screen "D_GraphicView_1" 800x480
   GraphicView "Static" at 6,4 size 100x60
   TextField "Label_Static" at 6,96 size 44x17; Text 'Static'
   GraphicView "A_Range" at 158,4 size 100x60
      Appearance <- "D_Range"
   TextField "Label_A_Range" at 158,96 size 63x17; Text 'A_Range'
   GraphicView "A_Flash" at 310,4 size 100x60
      Appearance <- "D_Range"
   TextField "Label_A_Flash" at 310,96 size 56x17; Text 'A_Flash'
   GraphicView "A_Bit" at 462,4 size 100x60
      Appearance <- "D_Bool"
   TextField "Label_A_Bit" at 462,96 size 40x17; Text 'A_Bit'
   GraphicView "A_Bits" at 614,4 size 100x60
      Appearance <- "D_Bits"
   TextField "Label_A_Bits" at 614,96 size 47x17; Text 'A_Bits'
   GraphicView "V_Range" at 6,116 size 100x60
      Visibility <- "D_Range"
   TextField "Label_V_Range" at 6,208 size 62x17; Text 'V_Range'
   GraphicView "V_Bit" at 158,116 size 100x60
      Visibility <- "D_Vis"
   TextField "Label_V_Bit" at 158,208 size 39x17; Text 'V_Bit'
   GraphicView "M_H" at 310,116 size 100x60
      HorizontalMovement <- "D_Pct"
   TextField "Label_M_H" at 310,208 size 33x17; Text 'M_H'
   GraphicView "M_V" at 462,116 size 100x60
      VerticalMovement <- "D_Pct"
   TextField "Label_M_V" at 462,208 size 32x17; Text 'M_V'
   GraphicView "M_D" at 614,116 size 100x60
      DiagonalMovement <- "D_Pct"
   TextField "Label_M_D" at 614,208 size 33x17; Text 'M_D'
   GraphicView "M_Direct" at 6,228 size 100x60
      DirectMovement <- "D_X"
      DirectMovement <- "D_Y"
   TextField "Label_M_Direct" at 6,320 size 64x17; Text 'M_Direct'
   GraphicView "E_Range" at 158,228 size 100x60
      ObjectEnable <- "D_Range"
   TextField "Label_E_Range" at 158,320 size 61x17; Text 'E_Range'
   GraphicView "E_Bit" at 310,228 size 100x60
      ObjectEnable <- "D_En"
   TextField "Label_E_Bit" at 310,320 size 38x17; Text 'E_Bit'
   IOField "State" at 4,454 size 60x22; FormatPattern 9
      ProcessValue <- "D_State"
   Button "S1" at 70,454 size 40x22; TextOff 'S1'
      on Click: "SetS1"()
   Button "S2" at 114,454 size 40x22; TextOff 'S2'
      on Click: "SetS2"()
   Button "S3" at 158,454 size 40x22; TextOff 'S3'
      on Click: "SetS3"()
   Button "S4" at 202,454 size 40x22; TextOff 'S4'
      on Click: "SetS4"()
   Button "Next" at 756,454 size 40x22; TextOff 'Next'
      on Click: ActivateScreen("D_IOField_1", 0)

screen "D_IOField_2" 800x480
   IOField "PV_Int_Output" at 6,4 size 100x30; FormatPattern s99999
      ProcessValue <- "D_Int"
   TextField "Label_PV_Int_Output" at 6,66 size 102x17; Text 'PV_Int_Output'
   IOField "PV_Int_s99" at 158,4 size 100x30; FormatPattern s99
      ProcessValue <- "D_Int"
   TextField "Label_PV_Int_s99" at 158,66 size 80x17; Text 'PV_Int_s99'
   IOField "State" at 4,454 size 60x22; FormatPattern 9
      ProcessValue <- "D_State"
   Button "S1" at 70,454 size 40x22; TextOff 'S1'
      on Click: "SetS1"()
   Button "S2" at 114,454 size 40x22; TextOff 'S2'
      on Click: "SetS2"()
   Button "S3" at 158,454 size 40x22; TextOff 'S3'
      on Click: "SetS3"()
   Button "S4" at 202,454 size 40x22; TextOff 'S4'
      on Click: "SetS4"()
   Button "Next" at 756,454 size 40x22; TextOff 'Next'
      on Click: ActivateScreen("D_Button_1", 0)

screen "D_Line_1" 800x480
   TextField "Label_Static" at 6,86 size 44x17; Text 'Static'
   Line "A_Range" at 158,4 size 100x50
      Appearance <- "D_Range"
   TextField "Label_A_Range" at 158,86 size 63x17; Text 'A_Range'
   Line "A_Flash" at 310,4 size 100x50
      Appearance <- "D_Range"
   TextField "Label_A_Flash" at 310,86 size 56x17; Text 'A_Flash'
   Line "A_Bit" at 462,4 size 100x50
      Appearance <- "D_Bool"
   TextField "Label_A_Bit" at 462,86 size 40x17; Text 'A_Bit'
   Line "A_Bits" at 614,4 size 100x50
      Appearance <- "D_Bits"
   TextField "Label_A_Bits" at 614,86 size 47x17; Text 'A_Bits'
   Line "V_Range" at 6,106 size 100x50
      Visibility <- "D_Range"
   TextField "Label_V_Range" at 6,188 size 62x17; Text 'V_Range'
   Line "V_Bit" at 158,106 size 100x50
      Visibility <- "D_Vis"
   TextField "Label_V_Bit" at 158,188 size 39x17; Text 'V_Bit'
   Line "M_H" at 310,106 size 100x50
      HorizontalMovement <- "D_Pct"
   TextField "Label_M_H" at 310,188 size 33x17; Text 'M_H'
   Line "M_V" at 462,106 size 100x50
      VerticalMovement <- "D_Pct"
   TextField "Label_M_V" at 462,188 size 32x17; Text 'M_V'
   Line "M_D" at 614,106 size 100x50
      DiagonalMovement <- "D_Pct"
   TextField "Label_M_D" at 614,188 size 33x17; Text 'M_D'
   Line "M_Direct" at 6,208 size 100x50
      DirectMovement <- "D_X"
      DirectMovement <- "D_Y"
   TextField "Label_M_Direct" at 6,290 size 64x17; Text 'M_Direct'
   Line "E_Range" at 158,208 size 100x50
      ObjectEnable <- "D_Range"
   TextField "Label_E_Range" at 158,290 size 61x17; Text 'E_Range'
   Line "E_Bit" at 310,208 size 100x50
      ObjectEnable <- "D_En"
   TextField "Label_E_Bit" at 310,290 size 38x17; Text 'E_Bit'
   IOField "State" at 4,454 size 60x22; FormatPattern 9
      ProcessValue <- "D_State"
   Button "S1" at 70,454 size 40x22; TextOff 'S1'
      on Click: "SetS1"()
   Button "S2" at 114,454 size 40x22; TextOff 'S2'
      on Click: "SetS2"()
   Button "S3" at 158,454 size 40x22; TextOff 'S3'
      on Click: "SetS3"()
   Button "S4" at 202,454 size 40x22; TextOff 'S4'
      on Click: "SetS4"()
   Button "Next" at 756,454 size 40x22; TextOff 'Next'
      on Click: ActivateScreen("D_Polyline_1", 0)

screen "D_Polygon_1" 800x480
   TextField "Label_Static" at 6,86 size 44x17; Text 'Static'
   Polygon "A_Range" at 158,4 size 100x50
      Appearance <- "D_Range"
   TextField "Label_A_Range" at 158,86 size 63x17; Text 'A_Range'
   Polygon "A_Flash" at 310,4 size 100x50
      Appearance <- "D_Range"
   TextField "Label_A_Flash" at 310,86 size 56x17; Text 'A_Flash'
   Polygon "A_Bit" at 462,4 size 100x50
      Appearance <- "D_Bool"
   TextField "Label_A_Bit" at 462,86 size 40x17; Text 'A_Bit'
   Polygon "A_Bits" at 614,4 size 100x50
      Appearance <- "D_Bits"
   TextField "Label_A_Bits" at 614,86 size 47x17; Text 'A_Bits'
   Polygon "V_Range" at 6,106 size 100x50
      Visibility <- "D_Range"
   TextField "Label_V_Range" at 6,188 size 62x17; Text 'V_Range'
   Polygon "V_Bit" at 158,106 size 100x50
      Visibility <- "D_Vis"
   TextField "Label_V_Bit" at 158,188 size 39x17; Text 'V_Bit'
   Polygon "M_H" at 310,106 size 100x50
      HorizontalMovement <- "D_Pct"
   TextField "Label_M_H" at 310,188 size 33x17; Text 'M_H'
   Polygon "M_V" at 462,106 size 100x50
      VerticalMovement <- "D_Pct"
   TextField "Label_M_V" at 462,188 size 32x17; Text 'M_V'
   Polygon "M_D" at 614,106 size 100x50
      DiagonalMovement <- "D_Pct"
   TextField "Label_M_D" at 614,188 size 33x17; Text 'M_D'
   Polygon "M_Direct" at 6,208 size 100x50
      DirectMovement <- "D_X"
      DirectMovement <- "D_Y"
   TextField "Label_M_Direct" at 6,290 size 64x17; Text 'M_Direct'
   Polygon "E_Range" at 158,208 size 100x50
      ObjectEnable <- "D_Range"
   TextField "Label_E_Range" at 158,290 size 61x17; Text 'E_Range'
   Polygon "E_Bit" at 310,208 size 100x50
      ObjectEnable <- "D_En"
   TextField "Label_E_Bit" at 310,290 size 38x17; Text 'E_Bit'
   IOField "State" at 4,454 size 60x22; FormatPattern 9
      ProcessValue <- "D_State"
   Button "S1" at 70,454 size 40x22; TextOff 'S1'
      on Click: "SetS1"()
   Button "S2" at 114,454 size 40x22; TextOff 'S2'
      on Click: "SetS2"()
   Button "S3" at 158,454 size 40x22; TextOff 'S3'
      on Click: "SetS3"()
   Button "S4" at 202,454 size 40x22; TextOff 'S4'
      on Click: "SetS4"()
   Button "Next" at 756,454 size 40x22; TextOff 'Next'
      on Click: ActivateScreen("D_Ellipse_1", 0)

screen "D_Polyline_1" 800x480
   TextField "Label_Static" at 6,86 size 44x17; Text 'Static'
   Polyline "A_Range" at 158,4 size 100x50
      Appearance <- "D_Range"
   TextField "Label_A_Range" at 158,86 size 63x17; Text 'A_Range'
   Polyline "A_Flash" at 310,4 size 100x50
      Appearance <- "D_Range"
   TextField "Label_A_Flash" at 310,86 size 56x17; Text 'A_Flash'
   Polyline "A_Bit" at 462,4 size 100x50
      Appearance <- "D_Bool"
   TextField "Label_A_Bit" at 462,86 size 40x17; Text 'A_Bit'
   Polyline "A_Bits" at 614,4 size 100x50
      Appearance <- "D_Bits"
   TextField "Label_A_Bits" at 614,86 size 47x17; Text 'A_Bits'
   Polyline "V_Range" at 6,106 size 100x50
      Visibility <- "D_Range"
   TextField "Label_V_Range" at 6,188 size 62x17; Text 'V_Range'
   Polyline "V_Bit" at 158,106 size 100x50
      Visibility <- "D_Vis"
   TextField "Label_V_Bit" at 158,188 size 39x17; Text 'V_Bit'
   Polyline "M_H" at 310,106 size 100x50
      HorizontalMovement <- "D_Pct"
   TextField "Label_M_H" at 310,188 size 33x17; Text 'M_H'
   Polyline "M_V" at 462,106 size 100x50
      VerticalMovement <- "D_Pct"
   TextField "Label_M_V" at 462,188 size 32x17; Text 'M_V'
   Polyline "M_D" at 614,106 size 100x50
      DiagonalMovement <- "D_Pct"
   TextField "Label_M_D" at 614,188 size 33x17; Text 'M_D'
   Polyline "M_Direct" at 6,208 size 100x50
      DirectMovement <- "D_X"
      DirectMovement <- "D_Y"
   TextField "Label_M_Direct" at 6,290 size 64x17; Text 'M_Direct'
   Polyline "E_Range" at 158,208 size 100x50
      ObjectEnable <- "D_Range"
   TextField "Label_E_Range" at 158,290 size 61x17; Text 'E_Range'
   Polyline "E_Bit" at 310,208 size 100x50
      ObjectEnable <- "D_En"
   TextField "Label_E_Bit" at 310,290 size 38x17; Text 'E_Bit'
   IOField "State" at 4,454 size 60x22; FormatPattern 9
      ProcessValue <- "D_State"
   Button "S1" at 70,454 size 40x22; TextOff 'S1'
      on Click: "SetS1"()
   Button "S2" at 114,454 size 40x22; TextOff 'S2'
      on Click: "SetS2"()
   Button "S3" at 158,454 size 40x22; TextOff 'S3'
      on Click: "SetS3"()
   Button "S4" at 202,454 size 40x22; TextOff 'S4'
      on Click: "SetS4"()
   Button "Next" at 756,454 size 40x22; TextOff 'Next'
      on Click: ActivateScreen("D_Polygon_1", 0)

screen "D_Rectangle_1" 800x480
   TextField "Label_Static" at 6,86 size 44x17; Text 'Static'
   Rectangle "A_Range" at 158,4 size 100x50
      Appearance <- "D_Range"
   TextField "Label_A_Range" at 158,86 size 63x17; Text 'A_Range'
   Rectangle "A_Flash" at 310,4 size 100x50
      Appearance <- "D_Range"
   TextField "Label_A_Flash" at 310,86 size 56x17; Text 'A_Flash'
   Rectangle "A_Bit" at 462,4 size 100x50
      Appearance <- "D_Bool"
   TextField "Label_A_Bit" at 462,86 size 40x17; Text 'A_Bit'
   Rectangle "A_Bits" at 614,4 size 100x50
      Appearance <- "D_Bits"
   TextField "Label_A_Bits" at 614,86 size 47x17; Text 'A_Bits'
   Rectangle "V_Range" at 6,106 size 100x50
      Visibility <- "D_Range"
   TextField "Label_V_Range" at 6,188 size 62x17; Text 'V_Range'
   Rectangle "V_Bit" at 158,106 size 100x50
      Visibility <- "D_Vis"
   TextField "Label_V_Bit" at 158,188 size 39x17; Text 'V_Bit'
   Rectangle "M_H" at 310,106 size 100x50
      HorizontalMovement <- "D_Pct"
   TextField "Label_M_H" at 310,188 size 33x17; Text 'M_H'
   Rectangle "M_V" at 462,106 size 100x50
      VerticalMovement <- "D_Pct"
   TextField "Label_M_V" at 462,188 size 32x17; Text 'M_V'
   Rectangle "M_D" at 614,106 size 100x50
      DiagonalMovement <- "D_Pct"
   TextField "Label_M_D" at 614,188 size 33x17; Text 'M_D'
   Rectangle "M_Direct" at 6,208 size 100x50
      DirectMovement <- "D_X"
      DirectMovement <- "D_Y"
   TextField "Label_M_Direct" at 6,290 size 64x17; Text 'M_Direct'
   Rectangle "E_Range" at 158,208 size 100x50
      ObjectEnable <- "D_Range"
   TextField "Label_E_Range" at 158,290 size 61x17; Text 'E_Range'
   Rectangle "E_Bit" at 310,208 size 100x50
      ObjectEnable <- "D_En"
   TextField "Label_E_Bit" at 310,290 size 38x17; Text 'E_Bit'
   IOField "State" at 4,454 size 60x22; FormatPattern 9
      ProcessValue <- "D_State"
   Button "S1" at 70,454 size 40x22; TextOff 'S1'
      on Click: "SetS1"()
   Button "S2" at 114,454 size 40x22; TextOff 'S2'
      on Click: "SetS2"()
   Button "S3" at 158,454 size 40x22; TextOff 'S3'
      on Click: "SetS3"()
   Button "S4" at 202,454 size 40x22; TextOff 'S4'
      on Click: "SetS4"()
   Button "Next" at 756,454 size 40x22; TextOff 'Next'
      on Click: ActivateScreen("D_TextField_1", 0)

screen "D_Switch_1" 800x480
   Switch "Static" at 6,4 size 120x40; CaptionText 'Switch'; TextOff '0'; TextOn '1'
   TextField "Label_Static" at 6,76 size 44x17; Text 'Static'
   Switch "A_Range" at 178,4 size 120x40; CaptionText 'Switch'; TextOff '0'; TextOn '1'
      Appearance <- "D_Range"
   TextField "Label_A_Range" at 178,76 size 63x17; Text 'A_Range'
   Switch "A_Flash" at 350,4 size 120x40; CaptionText 'Switch'; TextOff '0'; TextOn '1'
      Appearance <- "D_Range"
   TextField "Label_A_Flash" at 350,76 size 56x17; Text 'A_Flash'
   Switch "A_Bit" at 522,4 size 120x40; CaptionText 'Switch'; TextOff '0'; TextOn '1'
      Appearance <- "D_Bool"
   TextField "Label_A_Bit" at 522,76 size 40x17; Text 'A_Bit'
   Switch "A_Bits" at 6,96 size 120x40; CaptionText 'Switch'; TextOff '0'; TextOn '1'
      Appearance <- "D_Bits"
   TextField "Label_A_Bits" at 6,168 size 47x17; Text 'A_Bits'
   Switch "V_Range" at 178,96 size 120x40; CaptionText 'Switch'; TextOff '0'; TextOn '1'
      Visibility <- "D_Range"
   TextField "Label_V_Range" at 178,168 size 62x17; Text 'V_Range'
   Switch "V_Bit" at 350,96 size 120x40; CaptionText 'Switch'; TextOff '0'; TextOn '1'
      Visibility <- "D_Vis"
   TextField "Label_V_Bit" at 350,168 size 39x17; Text 'V_Bit'
   Switch "M_H" at 522,96 size 120x40; CaptionText 'Switch'; TextOff '0'; TextOn '1'
      HorizontalMovement <- "D_Pct"
   TextField "Label_M_H" at 522,168 size 33x17; Text 'M_H'
   Switch "M_V" at 6,188 size 120x40; CaptionText 'Switch'; TextOff '0'; TextOn '1'
      VerticalMovement <- "D_Pct"
   TextField "Label_M_V" at 6,260 size 32x17; Text 'M_V'
   Switch "M_D" at 178,188 size 120x40; CaptionText 'Switch'; TextOff '0'; TextOn '1'
      DiagonalMovement <- "D_Pct"
   TextField "Label_M_D" at 178,260 size 33x17; Text 'M_D'
   Switch "M_Direct" at 350,188 size 120x40; CaptionText 'Switch'; TextOff '0'; TextOn '1'
      DirectMovement <- "D_X"
      DirectMovement <- "D_Y"
   TextField "Label_M_Direct" at 350,260 size 64x17; Text 'M_Direct'
   Switch "E_Range" at 522,188 size 120x40; CaptionText 'Switch'; TextOff '0'; TextOn '1'
      ObjectEnable <- "D_Range"
   TextField "Label_E_Range" at 522,260 size 61x17; Text 'E_Range'
   Switch "E_Bit" at 6,280 size 120x40; CaptionText 'Switch'; TextOff '0'; TextOn '1'
      ObjectEnable <- "D_En"
   TextField "Label_E_Bit" at 6,352 size 38x17; Text 'E_Bit'
   Switch "PV_Bool" at 178,280 size 120x40; CaptionText 'Switch'; TextOff '0'; TextOn '1'
      ProcessValue <- "D_Bool"
   TextField "Label_PV_Bool" at 178,352 size 57x17; Text 'PV_Bool'
   IOField "State" at 4,454 size 60x22; FormatPattern 9
      ProcessValue <- "D_State"
   Button "S1" at 70,454 size 40x22; TextOff 'S1'
      on Click: "SetS1"()
   Button "S2" at 114,454 size 40x22; TextOff 'S2'
      on Click: "SetS2"()
   Button "S3" at 158,454 size 40x22; TextOff 'S3'
      on Click: "SetS3"()
   Button "S4" at 202,454 size 40x22; TextOff 'S4'
      on Click: "SetS4"()
   Button "Next" at 756,454 size 40x22; TextOff 'Next'
      on Click: ActivateScreen("D_SymbolLibrary_1", 0)

screen "D_SymbolicIOField_1" 800x480
   SymbolicIOField "Static" at 6,4 size 120x30; TextOff '0'; TextOn '1'
   TextField "Label_Static" at 6,66 size 44x17; Text 'Static'
   SymbolicIOField "A_Range" at 178,4 size 120x30; TextOff '0'; TextOn '1'
      Appearance <- "D_Range"
   TextField "Label_A_Range" at 178,66 size 63x17; Text 'A_Range'
   SymbolicIOField "A_Flash" at 350,4 size 120x30; TextOff '0'; TextOn '1'
      Appearance <- "D_Range"
   TextField "Label_A_Flash" at 350,66 size 56x17; Text 'A_Flash'
   SymbolicIOField "A_Bit" at 522,4 size 120x30; TextOff '0'; TextOn '1'
      Appearance <- "D_Bool"
   TextField "Label_A_Bit" at 522,66 size 40x17; Text 'A_Bit'
   SymbolicIOField "A_Bits" at 6,86 size 120x30; TextOff '0'; TextOn '1'
      Appearance <- "D_Bits"
   TextField "Label_A_Bits" at 6,148 size 47x17; Text 'A_Bits'
   SymbolicIOField "V_Range" at 178,86 size 120x30; TextOff '0'; TextOn '1'
      Visibility <- "D_Range"
   TextField "Label_V_Range" at 178,148 size 62x17; Text 'V_Range'
   SymbolicIOField "V_Bit" at 350,86 size 120x30; TextOff '0'; TextOn '1'
      Visibility <- "D_Vis"
   TextField "Label_V_Bit" at 350,148 size 39x17; Text 'V_Bit'
   SymbolicIOField "M_H" at 522,86 size 120x30; TextOff '0'; TextOn '1'
      HorizontalMovement <- "D_Pct"
   TextField "Label_M_H" at 522,148 size 33x17; Text 'M_H'
   SymbolicIOField "M_V" at 6,168 size 120x30; TextOff '0'; TextOn '1'
      VerticalMovement <- "D_Pct"
   TextField "Label_M_V" at 6,230 size 32x17; Text 'M_V'
   SymbolicIOField "M_D" at 178,168 size 120x30; TextOff '0'; TextOn '1'
      DiagonalMovement <- "D_Pct"
   TextField "Label_M_D" at 178,230 size 33x17; Text 'M_D'
   SymbolicIOField "M_Direct" at 350,168 size 120x30; TextOff '0'; TextOn '1'
      DirectMovement <- "D_X"
      DirectMovement <- "D_Y"
   TextField "Label_M_Direct" at 350,230 size 64x17; Text 'M_Direct'
   SymbolicIOField "E_Range" at 522,168 size 120x30; TextOff '0'; TextOn '1'
      ObjectEnable <- "D_Range"
   TextField "Label_E_Range" at 522,230 size 61x17; Text 'E_Range'
   SymbolicIOField "E_Bit" at 6,250 size 120x30; TextOff '0'; TextOn '1'
      ObjectEnable <- "D_En"
   TextField "Label_E_Bit" at 6,312 size 38x17; Text 'E_Bit'
   SymbolicIOField "PV_TL_Value" at 178,250 size 120x30; TextOff '0'; TextOn '1'; TextList "TL_Value"
      ProcessValue <- "D_TL"
   TextField "Label_PV_TL_Value" at 178,312 size 88x17; Text 'PV_TL_Value'
   SymbolicIOField "PV_TL_Bit" at 350,250 size 120x30; TextOff '0'; TextOn '1'; TextList "TL_Bit"
      ProcessValue <- "D_Bool"
   TextField "Label_PV_TL_Bit" at 350,312 size 70x17; Text 'PV_TL_Bit'
   SymbolicIOField "PV_TL_BitNo" at 522,250 size 120x30; TextOff '0'; TextOn '1'; TextList "TL_BitNo"
      ProcessValue <- "D_Bits"
   TextField "Label_PV_TL_BitNo" at 522,312 size 86x17; Text 'PV_TL_BitNo'
   IOField "State" at 4,454 size 60x22; FormatPattern 9
      ProcessValue <- "D_State"
   Button "S1" at 70,454 size 40x22; TextOff 'S1'
      on Click: "SetS1"()
   Button "S2" at 114,454 size 40x22; TextOff 'S2'
      on Click: "SetS2"()
   Button "S3" at 158,454 size 40x22; TextOff 'S3'
      on Click: "SetS3"()
   Button "S4" at 202,454 size 40x22; TextOff 'S4'
      on Click: "SetS4"()
   Button "Next" at 756,454 size 40x22; TextOff 'Next'
      on Click: ActivateScreen("D_GraphicIOField_1", 0)

screen "D_TextField_1" 800x480
   TextField "Static" at 6,4 size 35x17; Text 'Text'
   TextField "Label_Static" at 6,66 size 44x17; Text 'Static'
   TextField "A_Range" at 158,4 size 35x17; Text 'Text'
      Appearance <- "D_Range"
   TextField "Label_A_Range" at 158,66 size 63x17; Text 'A_Range'
   TextField "A_Flash" at 310,4 size 35x17; Text 'Text'
      Appearance <- "D_Range"
   TextField "Label_A_Flash" at 310,66 size 56x17; Text 'A_Flash'
   TextField "A_Bit" at 462,4 size 35x17; Text 'Text'
      Appearance <- "D_Bool"
   TextField "Label_A_Bit" at 462,66 size 40x17; Text 'A_Bit'
   TextField "A_Bits" at 614,4 size 35x17; Text 'Text'
      Appearance <- "D_Bits"
   TextField "Label_A_Bits" at 614,66 size 47x17; Text 'A_Bits'
   TextField "V_Range" at 6,86 size 35x17; Text 'Text'
      Visibility <- "D_Range"
   TextField "Label_V_Range" at 6,148 size 62x17; Text 'V_Range'
   TextField "V_Bit" at 158,86 size 35x17; Text 'Text'
      Visibility <- "D_Vis"
   TextField "Label_V_Bit" at 158,148 size 39x17; Text 'V_Bit'
   TextField "M_H" at 310,86 size 35x17; Text 'Text'
      HorizontalMovement <- "D_Pct"
   TextField "Label_M_H" at 310,148 size 33x17; Text 'M_H'
   TextField "M_V" at 462,86 size 35x17; Text 'Text'
      VerticalMovement <- "D_Pct"
   TextField "Label_M_V" at 462,148 size 32x17; Text 'M_V'
   TextField "M_D" at 614,86 size 35x17; Text 'Text'
      DiagonalMovement <- "D_Pct"
   TextField "Label_M_D" at 614,148 size 33x17; Text 'M_D'
   TextField "M_Direct" at 6,168 size 35x17; Text 'Text'
      DirectMovement <- "D_X"
      DirectMovement <- "D_Y"
   TextField "Label_M_Direct" at 6,230 size 64x17; Text 'M_Direct'
   TextField "E_Range" at 158,168 size 35x17; Text 'Text'
      ObjectEnable <- "D_Range"
   TextField "Label_E_Range" at 158,230 size 61x17; Text 'E_Range'
   TextField "E_Bit" at 310,168 size 35x17; Text 'Text'
      ObjectEnable <- "D_En"
   TextField "Label_E_Bit" at 310,230 size 38x17; Text 'E_Bit'
   IOField "State" at 4,454 size 60x22; FormatPattern 9
      ProcessValue <- "D_State"
   Button "S1" at 70,454 size 40x22; TextOff 'S1'
      on Click: "SetS1"()
   Button "S2" at 114,454 size 40x22; TextOff 'S2'
      on Click: "SetS2"()
   Button "S3" at 158,454 size 40x22; TextOff 'S3'
      on Click: "SetS3"()
   Button "S4" at 202,454 size 40x22; TextOff 'S4'
      on Click: "SetS4"()
   Button "Next" at 756,454 size 40x22; TextOff 'Next'
      on Click: ActivateScreen("D_GraphicView_1", 0)

screen "D_IOField_1" 800x480
   IOField "Static" at 6,4 size 100x30
   TextField "Label_Static" at 6,66 size 44x17; Text 'Static'
   IOField "A_Range" at 158,4 size 100x30
      Appearance <- "D_Range"
   TextField "Label_A_Range" at 158,66 size 63x17; Text 'A_Range'
   IOField "A_Flash" at 310,4 size 100x30
      Appearance <- "D_Range"
   TextField "Label_A_Flash" at 310,66 size 56x17; Text 'A_Flash'
   IOField "A_Bit" at 462,4 size 100x30
      Appearance <- "D_Bool"
   TextField "Label_A_Bit" at 462,66 size 40x17; Text 'A_Bit'
   IOField "A_Bits" at 614,4 size 100x30
      Appearance <- "D_Bits"
   TextField "Label_A_Bits" at 614,66 size 47x17; Text 'A_Bits'
   IOField "V_Range" at 6,86 size 100x30
      Visibility <- "D_Range"
   TextField "Label_V_Range" at 6,148 size 62x17; Text 'V_Range'
   IOField "V_Bit" at 158,86 size 100x30
      Visibility <- "D_Vis"
   TextField "Label_V_Bit" at 158,148 size 39x17; Text 'V_Bit'
   IOField "M_H" at 310,86 size 100x30
      HorizontalMovement <- "D_Pct"
   TextField "Label_M_H" at 310,148 size 33x17; Text 'M_H'
   IOField "M_V" at 462,86 size 100x30
      VerticalMovement <- "D_Pct"
   TextField "Label_M_V" at 462,148 size 32x17; Text 'M_V'
   IOField "M_D" at 614,86 size 100x30
      DiagonalMovement <- "D_Pct"
   TextField "Label_M_D" at 614,148 size 33x17; Text 'M_D'
   IOField "M_Direct" at 6,168 size 100x30
      DirectMovement <- "D_X"
      DirectMovement <- "D_Y"
   TextField "Label_M_Direct" at 6,230 size 64x17; Text 'M_Direct'
   IOField "E_Range" at 158,168 size 100x30
      ObjectEnable <- "D_Range"
   TextField "Label_E_Range" at 158,230 size 61x17; Text 'E_Range'
   IOField "E_Bit" at 310,168 size 100x30
      ObjectEnable <- "D_En"
   TextField "Label_E_Bit" at 310,230 size 38x17; Text 'E_Bit'
   IOField "PV_SInt" at 462,168 size 100x30; FormatPattern s999
      ProcessValue <- "D_SInt"
   TextField "Label_PV_SInt" at 462,230 size 57x17; Text 'PV_SInt'
   IOField "PV_Int" at 614,168 size 100x30; FormatPattern s99999
      ProcessValue <- "D_Int"
   TextField "Label_PV_Int" at 614,230 size 49x17; Text 'PV_Int'
   IOField "PV_DInt" at 6,250 size 100x30; FormatPattern s9999999999
      ProcessValue <- "D_DInt"
   TextField "Label_PV_DInt" at 6,312 size 58x17; Text 'PV_DInt'
   IOField "PV_USInt" at 158,250 size 100x30; FormatPattern 999
      ProcessValue <- "D_USInt"
   TextField "Label_PV_USInt" at 158,312 size 66x17; Text 'PV_USInt'
   IOField "PV_UInt" at 310,250 size 100x30; FormatPattern 99999
      ProcessValue <- "D_UInt"
   TextField "Label_PV_UInt" at 310,312 size 58x17; Text 'PV_UInt'
   IOField "PV_UDInt" at 462,250 size 100x30; FormatPattern 9999999999
      ProcessValue <- "D_UDInt"
   TextField "Label_PV_UDInt" at 462,312 size 67x17; Text 'PV_UDInt'
   IOField "PV_Real" at 614,250 size 100x30
      ProcessValue <- "D_Real"
   TextField "Label_PV_Real" at 614,312 size 58x17; Text 'PV_Real'
   IOField "PV_LReal" at 6,332 size 100x30
      ProcessValue <- "D_LReal"
   TextField "Label_PV_LReal" at 6,394 size 65x17; Text 'PV_LReal'
   IOField "PV_String" at 158,332 size 100x30
      ProcessValue <- "D_String"
   TextField "Label_PV_String" at 158,394 size 69x17; Text 'PV_String'
   IOField "PV_Int_Shift2" at 310,332 size 100x30; FormatPattern s99999
      ProcessValue <- "D_Int"
   TextField "Label_PV_Int_Shift2" at 310,394 size 96x17; Text 'PV_Int_Shift2'
   IOField "PV_Int_s999999" at 462,332 size 100x30; FormatPattern s999999
      ProcessValue <- "D_Int"
   TextField "Label_PV_Int_s999999" at 462,394 size 112x17; Text 'PV_Int_s999999'
   IOField "PV_Real_s9999_99" at 614,332 size 100x30; FormatPattern s9999.99
      ProcessValue <- "D_Real"
   TextField "Label_PV_Real_s9999_99" at 614,394 size 129x17; Text 'PV_Real_s9999_99'
   IOField "State" at 4,454 size 60x22; FormatPattern 9
      ProcessValue <- "D_State"
   Button "S1" at 70,454 size 40x22; TextOff 'S1'
      on Click: "SetS1"()
   Button "S2" at 114,454 size 40x22; TextOff 'S2'
      on Click: "SetS2"()
   Button "S3" at 158,454 size 40x22; TextOff 'S3'
      on Click: "SetS3"()
   Button "S4" at 202,454 size 40x22; TextOff 'S4'
      on Click: "SetS4"()
   Button "Next" at 756,454 size 40x22; TextOff 'Next'
      on Click: ActivateScreen("D_IOField_2", 0)

screen "D_Bar_1" 800x480
   Bar "Static" at 6,4 size 40x120
   TextField "Label_Static" at 6,156 size 44x17; Text 'Static'
   Bar "A_Range" at 98,4 size 40x120
      Appearance <- "D_Range"
   TextField "Label_A_Range" at 98,156 size 63x17; Text 'A_Range'
   Bar "A_Flash" at 190,4 size 40x120
      Appearance <- "D_Range"
   TextField "Label_A_Flash" at 190,156 size 56x17; Text 'A_Flash'
   Bar "A_Bit" at 282,4 size 40x120
      Appearance <- "D_Bool"
   TextField "Label_A_Bit" at 282,156 size 40x17; Text 'A_Bit'
   Bar "A_Bits" at 374,4 size 40x120
      Appearance <- "D_Bits"
   TextField "Label_A_Bits" at 374,156 size 47x17; Text 'A_Bits'
   Bar "V_Range" at 466,4 size 40x120
      Visibility <- "D_Range"
   TextField "Label_V_Range" at 466,156 size 62x17; Text 'V_Range'
   Bar "V_Bit" at 558,4 size 40x120
      Visibility <- "D_Vis"
   TextField "Label_V_Bit" at 558,156 size 39x17; Text 'V_Bit'
   Bar "M_H" at 650,4 size 40x120
      HorizontalMovement <- "D_Pct"
   TextField "Label_M_H" at 650,156 size 33x17; Text 'M_H'
   Bar "M_V" at 6,176 size 40x120
      VerticalMovement <- "D_Pct"
   TextField "Label_M_V" at 6,328 size 32x17; Text 'M_V'
   Bar "M_D" at 98,176 size 40x120
      DiagonalMovement <- "D_Pct"
   TextField "Label_M_D" at 98,328 size 33x17; Text 'M_D'
   Bar "M_Direct" at 190,176 size 40x120
      DirectMovement <- "D_X"
      DirectMovement <- "D_Y"
   TextField "Label_M_Direct" at 190,328 size 64x17; Text 'M_Direct'
   Bar "E_Range" at 282,176 size 40x120
      ObjectEnable <- "D_Range"
   TextField "Label_E_Range" at 282,328 size 61x17; Text 'E_Range'
   Bar "E_Bit" at 374,176 size 40x120
      ObjectEnable <- "D_En"
   TextField "Label_E_Bit" at 374,328 size 38x17; Text 'E_Bit'
   Bar "PV_Pct" at 466,176 size 40x120
      ProcessValue <- "D_Pct"
   TextField "Label_PV_Pct" at 466,328 size 50x17; Text 'PV_Pct'
   Bar "PV_Real" at 558,176 size 40x120
      ProcessValue <- "D_Real"
   TextField "Label_PV_Real" at 558,328 size 58x17; Text 'PV_Real'
   Bar "PV_BarR" at 650,176 size 40x120
      ProcessValue <- "D_BarR"
   TextField "Label_PV_BarR" at 650,328 size 60x17; Text 'PV_BarR'
   IOField "State" at 4,454 size 60x22; FormatPattern 9
      ProcessValue <- "D_State"
   Button "S1" at 70,454 size 40x22; TextOff 'S1'
      on Click: "SetS1"()
   Button "S2" at 114,454 size 40x22; TextOff 'S2'
      on Click: "SetS2"()
   Button "S3" at 158,454 size 40x22; TextOff 'S3'
      on Click: "SetS3"()
   Button "S4" at 202,454 size 40x22; TextOff 'S4'
      on Click: "SetS4"()
   Button "Next" at 756,454 size 40x22; TextOff 'Next'
      on Click: ActivateScreen("D_Bar_2", 0)

screen "D_Bar_2" 800x480
   Bar "PV_Pct_0_100" at 6,4 size 40x120; MinimumValue 0; MaximumValue 100
      ProcessValue <- "D_Pct"
   TextField "Label_PV_Pct_0_100" at 6,156 size 98x17; Text 'PV_Pct_0_100'
   Bar "PV_Pct_MaxMin" at 98,4 size 40x120
      ProcessValue <- "D_Pct"
      MaximumValue <- "D_Max"
      MinimumValue <- "D_Min"
   TextField "Label_PV_Pct_MaxMin" at 98,156 size 108x17; Text 'PV_Pct_MaxMin'
   IOField "State" at 4,454 size 60x22; FormatPattern 9
      ProcessValue <- "D_State"
   Button "S1" at 70,454 size 40x22; TextOff 'S1'
      on Click: "SetS1"()
   Button "S2" at 114,454 size 40x22; TextOff 'S2'
      on Click: "SetS2"()
   Button "S3" at 158,454 size 40x22; TextOff 'S3'
      on Click: "SetS3"()
   Button "S4" at 202,454 size 40x22; TextOff 'S4'
      on Click: "SetS4"()
   Button "Next" at 756,454 size 40x22; TextOff 'Next'
      on Click: ActivateScreen("D_Switch_1", 0)

screen "D_Gauge_1" 800x480
   Gauge "Static" at 6,4 size 150x150; CaptionText 'SIMATIC'
   TextField "Label_Static" at 6,186 size 44x17; Text 'Static'
   Gauge "A_Range" at 208,4 size 150x150; CaptionText 'SIMATIC'
      Appearance <- "D_Range"
   TextField "Label_A_Range" at 208,186 size 63x17; Text 'A_Range'
   Gauge "A_Flash" at 410,4 size 150x150; CaptionText 'SIMATIC'
      Appearance <- "D_Range"
   TextField "Label_A_Flash" at 410,186 size 56x17; Text 'A_Flash'
   Gauge "A_Bit" at 6,206 size 150x150; CaptionText 'SIMATIC'
      Appearance <- "D_Bool"
   TextField "Label_A_Bit" at 6,388 size 40x17; Text 'A_Bit'
   Gauge "A_Bits" at 208,206 size 150x150; CaptionText 'SIMATIC'
      Appearance <- "D_Bits"
   TextField "Label_A_Bits" at 208,388 size 47x17; Text 'A_Bits'
   Gauge "V_Range" at 410,206 size 150x150; CaptionText 'SIMATIC'
      Visibility <- "D_Range"
   TextField "Label_V_Range" at 410,388 size 62x17; Text 'V_Range'
   IOField "State" at 4,454 size 60x22; FormatPattern 9
      ProcessValue <- "D_State"
   Button "S1" at 70,454 size 40x22; TextOff 'S1'
      on Click: "SetS1"()
   Button "S2" at 114,454 size 40x22; TextOff 'S2'
      on Click: "SetS2"()
   Button "S3" at 158,454 size 40x22; TextOff 'S3'
      on Click: "SetS3"()
   Button "S4" at 202,454 size 40x22; TextOff 'S4'
      on Click: "SetS4"()
   Button "Next" at 756,454 size 40x22; TextOff 'Next'
      on Click: ActivateScreen("D_Gauge_2", 0)

screen "D_Gauge_2" 800x480
   Gauge "V_Bit" at 6,4 size 150x150; CaptionText 'SIMATIC'
      Visibility <- "D_Vis"
   TextField "Label_V_Bit" at 6,186 size 39x17; Text 'V_Bit'
   Gauge "M_H" at 208,4 size 150x150; CaptionText 'SIMATIC'
      HorizontalMovement <- "D_Pct"
   TextField "Label_M_H" at 208,186 size 33x17; Text 'M_H'
   Gauge "M_V" at 410,4 size 150x150; CaptionText 'SIMATIC'
      VerticalMovement <- "D_Pct"
   TextField "Label_M_V" at 410,186 size 32x17; Text 'M_V'
   Gauge "M_D" at 6,206 size 150x150; CaptionText 'SIMATIC'
      DiagonalMovement <- "D_Pct"
   TextField "Label_M_D" at 6,388 size 33x17; Text 'M_D'
   Gauge "M_Direct" at 208,206 size 150x150; CaptionText 'SIMATIC'
      DirectMovement <- "D_X"
      DirectMovement <- "D_Y"
   TextField "Label_M_Direct" at 208,388 size 64x17; Text 'M_Direct'
   Gauge "E_Range" at 410,206 size 150x150; CaptionText 'SIMATIC'
      ObjectEnable <- "D_Range"
   TextField "Label_E_Range" at 410,388 size 61x17; Text 'E_Range'
   IOField "State" at 4,454 size 60x22; FormatPattern 9
      ProcessValue <- "D_State"
   Button "S1" at 70,454 size 40x22; TextOff 'S1'
      on Click: "SetS1"()
   Button "S2" at 114,454 size 40x22; TextOff 'S2'
      on Click: "SetS2"()
   Button "S3" at 158,454 size 40x22; TextOff 'S3'
      on Click: "SetS3"()
   Button "S4" at 202,454 size 40x22; TextOff 'S4'
      on Click: "SetS4"()
   Button "Next" at 756,454 size 40x22; TextOff 'Next'
      on Click: ActivateScreen("D_Gauge_3", 0)

screen "D_Gauge_3" 800x480
   Gauge "E_Bit" at 6,4 size 150x150; CaptionText 'SIMATIC'
      ObjectEnable <- "D_En"
   TextField "Label_E_Bit" at 6,186 size 38x17; Text 'E_Bit'
   Gauge "PV_Pct" at 208,4 size 150x150; CaptionText 'SIMATIC'
      ProcessValue <- "D_Pct"
   TextField "Label_PV_Pct" at 208,186 size 50x17; Text 'PV_Pct'
   Gauge "PV_Real" at 410,4 size 150x150; CaptionText 'SIMATIC'
      ProcessValue <- "D_Real"
   TextField "Label_PV_Real" at 410,186 size 58x17; Text 'PV_Real'
   Gauge "PV_Pct_MaxMin" at 6,206 size 150x150; CaptionText 'SIMATIC'
      ProcessValue <- "D_Pct"
      MaximumValue <- "D_Max"
      MinimumValue <- "D_Min"
   TextField "Label_PV_Pct_MaxMin" at 6,388 size 108x17; Text 'PV_Pct_MaxMin'
   IOField "State" at 4,454 size 60x22; FormatPattern 9
      ProcessValue <- "D_State"
   Button "S1" at 70,454 size 40x22; TextOff 'S1'
      on Click: "SetS1"()
   Button "S2" at 114,454 size 40x22; TextOff 'S2'
      on Click: "SetS2"()
   Button "S3" at 158,454 size 40x22; TextOff 'S3'
      on Click: "SetS3"()
   Button "S4" at 202,454 size 40x22; TextOff 'S4'
      on Click: "SetS4"()
   Button "Next" at 756,454 size 40x22; TextOff 'Next'
      on Click: ActivateScreen("D_Clock_1", 0)

screen "D_Slider_1" 800x480
   Slider "Static" at 6,4 size 60x160; Caption 'SIMATIC'
   TextField "Label_Static" at 6,196 size 44x17; Text 'Static'
   Slider "A_Range" at 118,4 size 60x160; Caption 'SIMATIC'
      Appearance <- "D_Range"
   TextField "Label_A_Range" at 118,196 size 63x17; Text 'A_Range'
   Slider "A_Flash" at 230,4 size 60x160; Caption 'SIMATIC'
      Appearance <- "D_Range"
   TextField "Label_A_Flash" at 230,196 size 56x17; Text 'A_Flash'
   Slider "A_Bit" at 342,4 size 60x160; Caption 'SIMATIC'
      Appearance <- "D_Bool"
   TextField "Label_A_Bit" at 342,196 size 40x17; Text 'A_Bit'
   Slider "A_Bits" at 454,4 size 60x160; Caption 'SIMATIC'
      Appearance <- "D_Bits"
   TextField "Label_A_Bits" at 454,196 size 47x17; Text 'A_Bits'
   Slider "V_Range" at 566,4 size 60x160; Caption 'SIMATIC'
      Visibility <- "D_Range"
   TextField "Label_V_Range" at 566,196 size 62x17; Text 'V_Range'
   Slider "V_Bit" at 678,4 size 60x160; Caption 'SIMATIC'
      Visibility <- "D_Vis"
   TextField "Label_V_Bit" at 678,196 size 39x17; Text 'V_Bit'
   Slider "M_H" at 6,216 size 60x160; Caption 'SIMATIC'
      HorizontalMovement <- "D_Pct"
   TextField "Label_M_H" at 6,408 size 33x17; Text 'M_H'
   Slider "M_V" at 118,216 size 60x160; Caption 'SIMATIC'
      VerticalMovement <- "D_Pct"
   TextField "Label_M_V" at 118,408 size 32x17; Text 'M_V'
   Slider "M_D" at 230,216 size 60x160; Caption 'SIMATIC'
      DiagonalMovement <- "D_Pct"
   TextField "Label_M_D" at 230,408 size 33x17; Text 'M_D'
   Slider "M_Direct" at 342,216 size 60x160; Caption 'SIMATIC'
      DirectMovement <- "D_X"
      DirectMovement <- "D_Y"
   TextField "Label_M_Direct" at 342,408 size 64x17; Text 'M_Direct'
   Slider "E_Range" at 454,216 size 60x160; Caption 'SIMATIC'
      ObjectEnable <- "D_Range"
   TextField "Label_E_Range" at 454,408 size 61x17; Text 'E_Range'
   Slider "E_Bit" at 566,216 size 60x160; Caption 'SIMATIC'
      ObjectEnable <- "D_En"
   TextField "Label_E_Bit" at 566,408 size 38x17; Text 'E_Bit'
   Slider "PV_Pct" at 678,216 size 60x160; Caption 'SIMATIC'
      ProcessValue <- "D_Pct"
   TextField "Label_PV_Pct" at 678,408 size 50x17; Text 'PV_Pct'
   IOField "State" at 4,454 size 60x22; FormatPattern 9
      ProcessValue <- "D_State"
   Button "S1" at 70,454 size 40x22; TextOff 'S1'
      on Click: "SetS1"()
   Button "S2" at 114,454 size 40x22; TextOff 'S2'
      on Click: "SetS2"()
   Button "S3" at 158,454 size 40x22; TextOff 'S3'
      on Click: "SetS3"()
   Button "S4" at 202,454 size 40x22; TextOff 'S4'
      on Click: "SetS4"()
   Button "Next" at 756,454 size 40x22; TextOff 'Next'
      on Click: ActivateScreen("D_Slider_2", 0)

screen "D_Slider_2" 800x480
   Slider "PV_Int" at 6,4 size 60x160; Caption 'SIMATIC'
      ProcessValue <- "D_Int"
   TextField "Label_PV_Int" at 6,196 size 49x17; Text 'PV_Int'
   Slider "PV_Pct_0_200" at 118,4 size 60x160; Caption 'SIMATIC'
      ProcessValue <- "D_Pct"
   TextField "Label_PV_Pct_0_200" at 118,196 size 98x17; Text 'PV_Pct_0_200'
   IOField "State" at 4,454 size 60x22; FormatPattern 9
      ProcessValue <- "D_State"
   Button "S1" at 70,454 size 40x22; TextOff 'S1'
      on Click: "SetS1"()
   Button "S2" at 114,454 size 40x22; TextOff 'S2'
      on Click: "SetS2"()
   Button "S3" at 158,454 size 40x22; TextOff 'S3'
      on Click: "SetS3"()
   Button "S4" at 202,454 size 40x22; TextOff 'S4'
      on Click: "SetS4"()
   Button "Next" at 756,454 size 40x22; TextOff 'Next'
      on Click: ActivateScreen("D_Gauge_1", 0)

screen "D_SymbolLibrary_1" 800x480
   SymbolLibrary "Static" at 6,4 size 60x60
   TextField "Label_Static" at 6,96 size 44x17; Text 'Static'
   SymbolLibrary "A_Range" at 118,4 size 60x60
      Appearance <- "D_Range"
   TextField "Label_A_Range" at 118,96 size 63x17; Text 'A_Range'
   SymbolLibrary "A_Flash" at 230,4 size 60x60
      Appearance <- "D_Range"
   TextField "Label_A_Flash" at 230,96 size 56x17; Text 'A_Flash'
   SymbolLibrary "A_Bit" at 342,4 size 60x60
      Appearance <- "D_Bool"
   TextField "Label_A_Bit" at 342,96 size 40x17; Text 'A_Bit'
   SymbolLibrary "A_Bits" at 454,4 size 60x60
      Appearance <- "D_Bits"
   TextField "Label_A_Bits" at 454,96 size 47x17; Text 'A_Bits'
   SymbolLibrary "V_Range" at 566,4 size 60x60
      Visibility <- "D_Range"
   TextField "Label_V_Range" at 566,96 size 62x17; Text 'V_Range'
   SymbolLibrary "V_Bit" at 678,4 size 60x60
      Visibility <- "D_Vis"
   TextField "Label_V_Bit" at 678,96 size 39x17; Text 'V_Bit'
   SymbolLibrary "M_H" at 6,116 size 60x60
      HorizontalMovement <- "D_Pct"
   TextField "Label_M_H" at 6,208 size 33x17; Text 'M_H'
   SymbolLibrary "M_V" at 118,116 size 60x60
      VerticalMovement <- "D_Pct"
   TextField "Label_M_V" at 118,208 size 32x17; Text 'M_V'
   SymbolLibrary "M_D" at 230,116 size 60x60
      DiagonalMovement <- "D_Pct"
   TextField "Label_M_D" at 230,208 size 33x17; Text 'M_D'
   SymbolLibrary "M_Direct" at 342,116 size 60x60
      DirectMovement <- "D_X"
      DirectMovement <- "D_Y"
   TextField "Label_M_Direct" at 342,208 size 64x17; Text 'M_Direct'
   SymbolLibrary "E_Range" at 454,116 size 60x60
      ObjectEnable <- "D_Range"
   TextField "Label_E_Range" at 454,208 size 61x17; Text 'E_Range'
   SymbolLibrary "E_Bit" at 566,116 size 60x60
      ObjectEnable <- "D_En"
   TextField "Label_E_Bit" at 566,208 size 38x17; Text 'E_Bit'
   SymbolLibrary "PV_Pct" at 678,116 size 60x60
      ProcessValue <- "D_Pct"
   TextField "Label_PV_Pct" at 678,208 size 50x17; Text 'PV_Pct'
   IOField "State" at 4,454 size 60x22; FormatPattern 9
      ProcessValue <- "D_State"
   Button "S1" at 70,454 size 40x22; TextOff 'S1'
      on Click: "SetS1"()
   Button "S2" at 114,454 size 40x22; TextOff 'S2'
      on Click: "SetS2"()
   Button "S3" at 158,454 size 40x22; TextOff 'S3'
      on Click: "SetS3"()
   Button "S4" at 202,454 size 40x22; TextOff 'S4'
      on Click: "SetS4"()
   Button "Next" at 756,454 size 40x22; TextOff 'Next'
      on Click: ActivateScreen("D_Slider_1", 0)

screen "C5_Buttons" 800x480, template "T_C05"
   Button "Btn_Text" at 6,40 size 120x50; TextOff 'Btn_Text off'; TextOn 'Btn_Text on'
   TextField "Label_Btn_Text" at 6,92 size 65x17; Text 'Btn_Text'
   Button "Btn_Graphic" at 182,40 size 120x90; TextOff 'Btn_Graphic off'; TextOn 'Btn_Graphic on'; PictureOff "G_PNG"; PictureOn "G_JPG"
   TextField "Label_Btn_Graphic" at 182,132 size 85x17; Text 'Btn_Graphic'
   Button "Btn_GraphicAndText" at 358,40 size 120x90; TextOff 'Btn_GraphicAndText off'; TextOn 'Btn_GraphicAndText on'; PictureOff "G_SVG"; PictureOn "G_EMF"
   TextField "Label_Btn_GraphicAndText" at 358,132 size 140x17; Text 'Btn_GraphicAndText'
   Button "Btn_TextList" at 534,40 size 160x50; TextOff 'Btn_TextList off'; TextOn 'Btn_TextList on'; TextList "TL_Value"
      ProcessValue <- "D_TL"
   TextField "Label_Btn_TextList" at 534,92 size 89x17; Text 'Btn_TextList'
   Button "Btn_GraphicList" at 6,152 size 120x90; TextOff 'Btn_GraphicList off'; TextOn 'Btn_GraphicList on'; PictureList "GL_Value"
      ProcessValue <- "D_TL"
   TextField "Label_Btn_GraphicList" at 6,244 size 109x17; Text 'Btn_GraphicList'
   Button "Btn_Invisible" at 182,152 size 120x50; TextOff 'Btn_Invisible off'; TextOn 'Btn_Invisible on'
   TextField "Label_Btn_Invisible" at 182,204 size 92x17; Text 'Btn_Invisible'
   Switch "Sw_Switch" at 358,152 size 120x40; CaptionText 'Switch'; TextOff '0'; TextOn '1'
      ProcessValue <- "D_Bool"
   TextField "Label_Sw_Switch" at 358,194 size 74x17; Text 'Sw_Switch'
   Switch "Sw_Text" at 534,152 size 120x40; CaptionText 'Switch'; TextOff 'Sw_Text off'; TextOn 'Sw_Text on'
      ProcessValue <- "D_Bool"
   TextField "Label_Sw_Text" at 534,194 size 61x17; Text 'Sw_Text'
   Switch "Sw_Graphic" at 6,264 size 120x90; CaptionText 'Switch'; TextOff '0'; TextOn '1'; PictureOff "G_BMP"; PictureOn "G_GIF"
      ProcessValue <- "D_Bool"
   TextField "Label_Sw_Graphic" at 6,356 size 81x17; Text 'Sw_Graphic'
   IOField "State" at 4,454 size 60x22; FormatPattern 9
      ProcessValue <- "D_State"
   Button "S1" at 70,454 size 40x22; TextOff 'S1'
      on Click: "SetS1"()
   Button "S2" at 114,454 size 40x22; TextOff 'S2'
      on Click: "SetS2"()
   Button "S3" at 158,454 size 40x22; TextOff 'S3'
      on Click: "SetS3"()
   Button "S4" at 202,454 size 40x22; TextOff 'S4'
      on Click: "SetS4"()
   Button "Next" at 756,454 size 40x22; TextOff 'Next'
      on Click: ActivateScreen("C5_Structure", 0)

screen "C5_GraphicView_1" 800x480, template "T_C05"
   GraphicView "GV_PNG" at 6,40 size 120x80; Picture "G_PNG"
   TextField "Label_GV_PNG" at 6,122 size 55x17; Text 'GV_PNG'
   GraphicView "GV_JPG" at 142,40 size 120x80; Picture "G_JPG"
   TextField "Label_GV_JPG" at 142,122 size 54x17; Text 'GV_JPG'
   GraphicView "GV_BMP" at 278,40 size 120x80; Picture "G_BMP"
   TextField "Label_GV_BMP" at 278,122 size 57x17; Text 'GV_BMP'
   GraphicView "GV_GIF" at 414,40 size 120x80; Picture "G_GIF"
   TextField "Label_GV_GIF" at 414,122 size 52x17; Text 'GV_GIF'
   GraphicView "GV_TIF" at 550,40 size 120x80; Picture "G_TIF"
   TextField "Label_GV_TIF" at 550,122 size 51x17; Text 'GV_TIF'
   GraphicView "GV_EMF" at 6,142 size 120x80; Picture "G_EMF"
   TextField "Label_GV_EMF" at 6,224 size 55x17; Text 'GV_EMF'
   GraphicView "GV_WMF" at 142,142 size 120x80; Picture "G_WMF"
   TextField "Label_GV_WMF" at 142,224 size 60x17; Text 'GV_WMF'
   GraphicView "GV_SVG" at 278,142 size 120x80; Picture "G_SVG"
   TextField "Label_GV_SVG" at 278,224 size 55x17; Text 'GV_SVG'
   GraphicView "GV_TALL" at 414,142 size 120x80; Picture "G_TALL"
   TextField "Label_GV_TALL" at 414,224 size 61x17; Text 'GV_TALL'
   GraphicView "GV_WIDE" at 550,142 size 120x80; Picture "G_WIDE"
   TextField "Label_GV_WIDE" at 550,224 size 64x17; Text 'GV_WIDE'
   IOField "State" at 4,454 size 60x22; FormatPattern 9
      ProcessValue <- "D_State"
   Button "S1" at 70,454 size 40x22; TextOff 'S1'
      on Click: "SetS1"()
   Button "S2" at 114,454 size 40x22; TextOff 'S2'
      on Click: "SetS2"()
   Button "S3" at 158,454 size 40x22; TextOff 'S3'
      on Click: "SetS3"()
   Button "S4" at 202,454 size 40x22; TextOff 'S4'
      on Click: "SetS4"()
   Button "Next" at 756,454 size 40x22; TextOff 'Next'
      on Click: ActivateScreen("C5_GraphicView_2_a", 0)

screen "C5_GraphicView_2_a" 800x480, template "T_C05"
   GraphicView "PNG_160x60_FitF" at 6,40 size 160x60; Picture "G_PNG"
   TextField "Label_PNG_160x60_FitF" at 6,102 size 118x17; Text 'PNG_160x60_FitF'
   GraphicView "PNG_160x60_FitT" at 182,40 size 160x60; Picture "G_PNG"
   TextField "Label_PNG_160x60_FitT" at 182,102 size 119x17; Text 'PNG_160x60_FitT'
   GraphicView "PNG_60x120_FitF" at 358,40 size 60x120; Picture "G_PNG"
   TextField "Label_PNG_60x120_FitF" at 358,162 size 118x17; Text 'PNG_60x120_FitF'
   GraphicView "PNG_60x120_FitT" at 534,40 size 60x120; Picture "G_PNG"
   TextField "Label_PNG_60x120_FitT" at 534,162 size 119x17; Text 'PNG_60x120_FitT'
   GraphicView "PNG_80x80_FitF" at 6,182 size 80x80; Picture "G_PNG"
   TextField "Label_PNG_80x80_FitF" at 6,264 size 110x17; Text 'PNG_80x80_FitF'
   GraphicView "PNG_80x80_FitT" at 182,182 size 80x80; Picture "G_PNG"
   TextField "Label_PNG_80x80_FitT" at 182,264 size 111x17; Text 'PNG_80x80_FitT'
   GraphicView "TALL_160x60_FitF" at 358,182 size 160x60; Picture "G_TALL"
   TextField "Label_TALL_160x60_FitF" at 358,244 size 124x17; Text 'TALL_160x60_FitF'
   GraphicView "TALL_160x60_FitT" at 534,182 size 160x60; Picture "G_TALL"
   TextField "Label_TALL_160x60_FitT" at 534,244 size 125x17; Text 'TALL_160x60_FitT'
   IOField "State" at 4,454 size 60x22; FormatPattern 9
      ProcessValue <- "D_State"
   Button "S1" at 70,454 size 40x22; TextOff 'S1'
      on Click: "SetS1"()
   Button "S2" at 114,454 size 40x22; TextOff 'S2'
      on Click: "SetS2"()
   Button "S3" at 158,454 size 40x22; TextOff 'S3'
      on Click: "SetS3"()
   Button "S4" at 202,454 size 40x22; TextOff 'S4'
      on Click: "SetS4"()
   Button "Next" at 756,454 size 40x22; TextOff 'Next'
      on Click: ActivateScreen("C5_GraphicView_2_b", 0)

screen "C5_GraphicView_2_b" 800x480, template "T_C05"
   GraphicView "TALL_60x120_FitF" at 6,40 size 60x120; Picture "G_TALL"
   TextField "Label_TALL_60x120_FitF" at 6,162 size 124x17; Text 'TALL_60x120_FitF'
   GraphicView "TALL_60x120_FitT" at 182,40 size 60x120; Picture "G_TALL"
   TextField "Label_TALL_60x120_FitT" at 182,162 size 125x17; Text 'TALL_60x120_FitT'
   GraphicView "TALL_80x80_FitF" at 358,40 size 80x80; Picture "G_TALL"
   TextField "Label_TALL_80x80_FitF" at 358,122 size 116x17; Text 'TALL_80x80_FitF'
   GraphicView "TALL_80x80_FitT" at 534,40 size 80x80; Picture "G_TALL"
   TextField "Label_TALL_80x80_FitT" at 534,122 size 117x17; Text 'TALL_80x80_FitT'
   GraphicView "WIDE_160x60_FitF" at 6,182 size 160x60; Picture "G_WIDE"
   TextField "Label_WIDE_160x60_FitF" at 6,244 size 127x17; Text 'WIDE_160x60_FitF'
   GraphicView "WIDE_160x60_FitT" at 182,182 size 160x60; Picture "G_WIDE"
   TextField "Label_WIDE_160x60_FitT" at 182,244 size 128x17; Text 'WIDE_160x60_FitT'
   GraphicView "WIDE_60x120_FitF" at 358,182 size 60x120; Picture "G_WIDE"
   TextField "Label_WIDE_60x120_FitF" at 358,304 size 127x17; Text 'WIDE_60x120_FitF'
   GraphicView "WIDE_60x120_FitT" at 534,182 size 60x120; Picture "G_WIDE"
   TextField "Label_WIDE_60x120_FitT" at 534,304 size 128x17; Text 'WIDE_60x120_FitT'
   IOField "State" at 4,454 size 60x22; FormatPattern 9
      ProcessValue <- "D_State"
   Button "S1" at 70,454 size 40x22; TextOff 'S1'
      on Click: "SetS1"()
   Button "S2" at 114,454 size 40x22; TextOff 'S2'
      on Click: "SetS2"()
   Button "S3" at 158,454 size 40x22; TextOff 'S3'
      on Click: "SetS3"()
   Button "S4" at 202,454 size 40x22; TextOff 'S4'
      on Click: "SetS4"()
   Button "Next" at 756,454 size 40x22; TextOff 'Next'
      on Click: ActivateScreen("C5_GraphicView_2_c", 0)

screen "C5_GraphicView_2_c" 800x480, template "T_C05"
   GraphicView "WIDE_80x80_FitF" at 6,40 size 80x80; Picture "G_WIDE"
   TextField "Label_WIDE_80x80_FitF" at 6,122 size 119x17; Text 'WIDE_80x80_FitF'
   GraphicView "WIDE_80x80_FitT" at 142,40 size 80x80; Picture "G_WIDE"
   TextField "Label_WIDE_80x80_FitT" at 142,122 size 120x17; Text 'WIDE_80x80_FitT'
   GraphicView "BMP_Transparent" at 278,40 size 120x80; Picture "G_BMP"
   TextField "Label_BMP_Transparent" at 278,122 size 121x17; Text 'BMP_Transparent'
   GraphicView "PNG_BackTransparent" at 414,40 size 120x80; Picture "G_PNG"
   TextField "Label_PNG_BackTransparent" at 414,122 size 150x17; Text 'PNG_BackTransparent'
   IOField "State" at 4,454 size 60x22; FormatPattern 9
      ProcessValue <- "D_State"
   Button "S1" at 70,454 size 40x22; TextOff 'S1'
      on Click: "SetS1"()
   Button "S2" at 114,454 size 40x22; TextOff 'S2'
      on Click: "SetS2"()
   Button "S3" at 158,454 size 40x22; TextOff 'S3'
      on Click: "SetS3"()
   Button "S4" at 202,454 size 40x22; TextOff 'S4'
      on Click: "SetS4"()
   Button "Next" at 756,454 size 40x22; TextOff 'Next'
      on Click: ActivateScreen("C5_Lists", 0)

screen "C5_Lists" 800x480, template "T_C05"
   SymbolicIOField "SIO_TL_Value" at 6,40 size 160x30; TextOff '0'; TextOn '1'; TextList "TL_Value"
      ProcessValue <- "D_TL"
   TextField "Label_SIO_TL_Value" at 6,72 size 95x17; Text 'SIO_TL_Value'
   SymbolicIOField "SIO_TL_Bit" at 182,40 size 160x30; TextOff '0'; TextOn '1'; TextList "TL_Bit"
      ProcessValue <- "D_Bool"
   TextField "Label_SIO_TL_Bit" at 182,72 size 77x17; Text 'SIO_TL_Bit'
   SymbolicIOField "SIO_TL_BitNo" at 358,40 size 160x30; TextOff '0'; TextOn '1'; TextList "TL_BitNo"
      ProcessValue <- "D_Bits"
   TextField "Label_SIO_TL_BitNo" at 358,72 size 93x17; Text 'SIO_TL_BitNo'
   SymbolicIOField "SIO_TL_Value_Out" at 534,40 size 160x30; TextOff '0'; TextOn '1'; TextList "TL_Value"
      ProcessValue <- "D_TL"
   TextField "Label_SIO_TL_Value_Out" at 534,72 size 126x17; Text 'SIO_TL_Value_Out'
   GraphicIOField "GIO_GL_Value" at 6,142 size 120x80; PictureList "GL_Value"
      ProcessValue <- "D_TL"
   TextField "Label_GIO_GL_Value" at 6,224 size 97x17; Text 'GIO_GL_Value'
   GraphicIOField "GIO_GL_Bit" at 182,142 size 120x80; PictureList "GL_Bit"
      ProcessValue <- "D_Bool"
   TextField "Label_GIO_GL_Bit" at 182,224 size 79x17; Text 'GIO_GL_Bit'
   GraphicIOField "GIO_GL_BitNo" at 358,142 size 120x80; PictureList "GL_BitNo"
      ProcessValue <- "D_Bits"
   TextField "Label_GIO_GL_BitNo" at 358,224 size 95x17; Text 'GIO_GL_BitNo'
   GraphicIOField "GIO_GL_Value_Out" at 534,142 size 120x80; PictureList "GL_Value"
      ProcessValue <- "D_TL"
   TextField "Label_GIO_GL_Value_Out" at 534,224 size 128x17; Text 'GIO_GL_Value_Out'
   IOField "State" at 4,454 size 60x22; FormatPattern 9
      ProcessValue <- "D_State"
   Button "S1" at 70,454 size 40x22; TextOff 'S1'
      on Click: "SetS1"()
   Button "S2" at 114,454 size 40x22; TextOff 'S2'
      on Click: "SetS2"()
   Button "S3" at 158,454 size 40x22; TextOff 'S3'
      on Click: "SetS3"()
   Button "S4" at 202,454 size 40x22; TextOff 'S4'
      on Click: "SetS4"()
   Button "Next" at 756,454 size 40x22; TextOff 'Next'
      on Click: ActivateScreen("C5_Buttons", 0)

Template "T_C05" 800x480
   TextField "T_Title" at 8,6 size 185x21; Text 'Template T_C05 (header)'
   DateTimeField "T_Clock" at 610,4 size 189x26

PopupScreen "Popup_C05" 300x200
   TextField "Pop_Title" at 10,10 size 175x17; Text 'Pop-up screen Popup_C05'
   GraphicView "Pop_Graphic" at 10,40 size 120x80; Picture "G_PNG"
   IOField "Pop_Value" at 150,60 size 120x30; FormatPattern s99999
      ProcessValue <- "D_Int"
   Button "Pop_Close" at 200,160 size 80x22; TextOff 'Close'
      on Click: function_efd93a16("Popup_C05", 200, 120, -1, -1, 1)

screen "C5_Structure" 800x480, template "T_C05"
   Group "Group_A" at 10,50 size 300x82
   TextField "Label_Group_A (contains Group_B)" at 10,140 size 192x17; Text 'Group_A (contains Group_B)'
   TextField "Layer0_Text" at 352,52 size 54x17; Text 'Layer 0'
   TextField "Label_Layers 0-3 (layer 2 VisibleES false)" at 350,200 size 235x17; Text 'Layers 0-3 (layer 2 VisibleES false)'
   IOField "State" at 4,454 size 60x22; FormatPattern 9
      ProcessValue <- "D_State"
   Button "S1" at 70,454 size 40x22; TextOff 'S1'
      on Click: "SetS1"()
   Button "S2" at 114,454 size 40x22; TextOff 'S2'
      on Click: "SetS2"()
   Button "S3" at 158,454 size 40x22; TextOff 'S3'
      on Click: "SetS3"()
   Button "S4" at 202,454 size 40x22; TextOff 'S4'
      on Click: "SetS4"()
   Button "Popup" at 246,454 size 60x22; TextOff 'Popup'
      on Click: function_efd93a16("Popup_C05", 200, 120, -1, -1, 1)
   Button "SlideIn" at 310,454 size 60x22; TextOff 'Slide'
      on Click: "C5_ToggleSlideIn"()
   Button "Next" at 756,454 size 40x22; TextOff 'Next'
      on Click: ActivateScreen("C5_GraphicView_1", 0)
   Group "Group_B" at 210,50 size 100x82
   TextField "GB_Text" at 210,115 size 60x17; Text 'Group_B'
   TextField "Layer1_Text" at 382,72 size 54x17; Text 'Layer 1'
   TextField "Layer2_Text" at 412,92 size 54x17; Text 'Layer 2'
   TextField "Layer3_Text" at 442,112 size 54x17; Text 'Layer 3'

screen "C6_Faceplates" 800x480
   ScreenModuleView "FP_Dyn" at 10,10 size 300x150; ScreenModuleType ""; Guid_{11997190-83750} 'Tags D_Int D_Range D_Pct'
      Guid_{11997190-83886} <- "D_Int"
      Guid_{11997190-83896} <- "D_Range"
      Guid_{11997190-83898} <- "D_Pct"
      Guid_{11997190-83900} <- "D_Vis"
   TextField "Label_FP_Dyn" at 10,162 size 53x17; Text 'FP_Dyn'
   ScreenModuleView "FP_Static" at 330,10 size 300x150; ScreenModuleType ""; Guid_{11997190-83750} 'Static values'
   TextField "Label_FP_Static" at 330,162 size 67x17; Text 'FP_Static'
   ScreenModuleView "FP_Alt" at 10,186 size 300x150; ScreenModuleType ""; Guid_{11997190-83750} 'Tags D_SInt D_TL D_UInt'
      Guid_{11997190-83886} <- "D_SInt"
      Guid_{11997190-83896} <- "D_TL"
      Guid_{11997190-83898} <- "D_UInt"
      Guid_{11997190-83900} <- "D_En"
   TextField "Label_FP_Alt" at 10,338 size 47x17; Text 'FP_Alt'
   ScreenModuleView "FP_Move" at 330,186 size 300x150; ScreenModuleType ""; Guid_{11997190-83750} 'Moved by D_Pct'
      Guid_{11997190-83886} <- "D_Int"
      Guid_{11997190-83896} <- "D_Range"
      Guid_{11997190-83898} <- "D_Pct"
      Guid_{11997190-83900} <- "D_Vis"
      HorizontalMovement <- "D_Pct"
   TextField "Label_FP_Move" at 330,338 size 63x17; Text 'FP_Move'
   IOField "State" at 4,454 size 60x22; FormatPattern 9
      ProcessValue <- "D_State"
   Button "S1" at 70,454 size 40x22; TextOff 'S1'
      on Click: "SetS1"()
   Button "S2" at 114,454 size 40x22; TextOff 'S2'
      on Click: "SetS2"()
   Button "S3" at 158,454 size 40x22; TextOff 'S3'
      on Click: "SetS3"()
   Button "S4" at 202,454 size 40x22; TextOff 'S4'
      on Click: "SetS4"()
   Button "Next" at 756,454 size 40x22; TextOff 'Next'
      on Click: ActivateScreen("C6_Faceplates", 0)

VB script "SetS1"
   SmartTags("D_State") = 1
   SmartTags("D_Bool") = False
   SmartTags("D_SInt") = -128
   SmartTags("D_Int") = -32768
   SmartTags("D_DInt") = -2147483648
   SmartTags("D_USInt") = 0
   SmartTags("D_UInt") = 0
   SmartTags("D_UDInt") = 0
   SmartTags("D_Real") = -999.999
   SmartTags("D_LReal") = -0.00000015
   SmartTags("D_String") = ""
   SmartTags("D_DateTime") = DateSerial(1990, 1, 1) + TimeSerial(0, 0, 0)
   SmartTags("D_Pct") = 0
   SmartTags("D_Range") = 5
   SmartTags("D_Bits") = 1
   SmartTags("D_Vis") = False
   SmartTags("D_En") = False
   SmartTags("D_X") = 10
   SmartTags("D_Y") = 10
   SmartTags("D_Max") = 100
   SmartTags("D_Min") = 0
   SmartTags("D_TL") = -5
   SmartTags("D_BarR") = -5

VB script "SetS2"
   SmartTags("D_State") = 2
   SmartTags("D_Bool") = True
   SmartTags("D_SInt") = 12
   SmartTags("D_Int") = 1234
   SmartTags("D_DInt") = 123456
   SmartTags("D_USInt") = 200
   SmartTags("D_UInt") = 40000
   SmartTags("D_UDInt") = 3000000000
   SmartTags("D_Real") = 3.14159
   SmartTags("D_LReal") = 2.718281828
   SmartTags("D_String") = "Hello World"
   SmartTags("D_DateTime") = DateSerial(2026, 11, 22) + TimeSerial(13, 45, 30)
   SmartTags("D_Pct") = 50
   SmartTags("D_Range") = 25
   SmartTags("D_Bits") = 2
   SmartTags("D_Vis") = True
   SmartTags("D_En") = True
   SmartTags("D_X") = 200
   SmartTags("D_Y") = 120
   SmartTags("D_Max") = 200
   SmartTags("D_Min") = -100
   SmartTags("D_TL") = 5
   SmartTags("D_BarR") = 0

VB script "SetS3"
   SmartTags("D_State") = 3
   SmartTags("D_Bool") = True
   SmartTags("D_SInt") = 127
   SmartTags("D_Int") = 32767
   SmartTags("D_DInt") = 2147483647
   SmartTags("D_USInt") = 255
   SmartTags("D_UInt") = 65535
   SmartTags("D_UDInt") = 4294967295
   SmartTags("D_Real") = 123456.789
   SmartTags("D_LReal") = 1E+300
   SmartTags("D_String") = "Ünïcödé äöüß ÄÖÜ € – long text that is wider than the field 0123456789 ABCDEFGHIJ"
   SmartTags("D_DateTime") = DateSerial(2099, 12, 31) + TimeSerial(23, 59, 59)
   SmartTags("D_Pct") = 100
   SmartTags("D_Range") = 75
   SmartTags("D_Bits") = 4
   SmartTags("D_Vis") = True
   SmartTags("D_En") = False
   SmartTags("D_X") = 533
   SmartTags("D_Y") = 240
   SmartTags("D_Max") = 50
   SmartTags("D_Min") = -50
   SmartTags("D_TL") = 10
   SmartTags("D_BarR") = 5

VB script "SetS4"
   SmartTags("D_State") = 4
   SmartTags("D_Bool") = False
   SmartTags("D_SInt") = -1
   SmartTags("D_Int") = -1
   SmartTags("D_DInt") = 0
   SmartTags("D_USInt") = 1
   SmartTags("D_UInt") = 1
   SmartTags("D_UDInt") = 1
   SmartTags("D_Real") = 0.0005
   SmartTags("D_LReal") = -0.0
   SmartTags("D_String") = "äöü ÄÖÜ ß"
   SmartTags("D_DateTime") = DateSerial(1970, 1, 1) + TimeSerial(0, 0, 0)
   SmartTags("D_Pct") = 150
   SmartTags("D_Range") = 200
   SmartTags("D_Bits") = 9
   SmartTags("D_Vis") = False
   SmartTags("D_En") = True
   SmartTags("D_X") = -20
   SmartTags("D_Y") = 0
   SmartTags("D_Max") = 100
   SmartTags("D_Min") = 0
   SmartTags("D_TL") = 50
   SmartTags("D_BarR") = 2.5

VB script "C5_ToggleSlideIn"
   cf6f4242-93bf-47b4-8281-e920249d00b8 GraphX_Slidein_Top, $3$hmiToggle$
*)

(* ===== HMI "HMI_RT_1" =====
system functions are stored by id; their names below are inferred from use
connection "HMI_Connection_3": ETHERNET, S7_1500_OMS

HMI tags "Default tag table"
   "Hmi_Bool" : Bool, internal
   "Hmi_Int" : Int, internal
   "Hmi_Real" : Real, internal
   "Hmi_String" : WString[254], internal
   "Ext_Bool" : Bool = PLC Plc_Bool AT %M100.0, 1 s
   "Ext_Int" : Int = PLC Plc_Int AT %MW102, 1 s
   "Ext_Real" : Real = PLC Plc_Real AT %MD104, 1 s
   "Ext_Byte" : Byte = PLC Plc_Byte AT %MB108, 1 s

HMI tags "C03_Tags"
   "D_State" : Int, internal
   "D_Bool" : Bool, internal
   "D_SInt" : SInt, internal
   "D_Int" : Int, internal
   "D_DInt" : DInt, internal
   "D_USInt" : USInt, internal
   "D_UInt" : UInt, internal
   "D_UDInt" : UDInt, internal
   "D_Real" : Real, internal
   "D_LReal" : LReal, internal
   "D_String" : WString[254], internal
   "D_DateTime" : DateTime, internal
   "D_Pct" : Int, internal
   "D_Range" : Int, internal
   "D_Bits" : Int, internal
   "D_Vis" : Bool, internal
   "D_En" : Bool, internal
   "D_X" : Int, internal
   "D_Y" : Int, internal
   "D_Max" : Real, internal
   "D_Min" : Real, internal
   "D_TL" : Int, internal
   "D_BarR" : Real, internal

discrete alarms
   1: 'Alarm bit 0 (D_Bits)', class Errors, trigger "D_Bits" bit 0
   2: 'Alarm bit 1 (D_Bits)', class Errors, trigger "D_Bits" bit 1
   3: 'Alarm bit 2 (D_Bits)', class Warnings, trigger "D_Bits" bit 2
   4: 'Alarm bit 3 (D_Bits)', class Warnings, trigger "D_Bits" bit 3

analog alarms
   1: 'D_Range above 50', class Errors, trigger "D_Range"

text list "TL_Bit": 0 'Off (0)'; 1 'On (1)'

text list "TL_BitNo": 0 'Bit 0 set'; 1 'Bit 1 set'; 2 'Bit 2 set'; 3 'Bit 3 set'

text list "TL_Value": -100..-1 'Negative (-100..-1)'; 0 'Zero'; 1..9 'One to nine'; 10 'Ten: Ünïcödé äöüß ÄÖÜ €'; 32000 'Undefined value (default entry)'

graphic list "GL_Bit": 0 'G_EMF'; 1 'G_WMF'

graphic list "GL_BitNo": 0 'G_PNG'; 1 'G_JPG'; 2 'G_BMP'; 3 'G_TIF'

graphic list "GL_Value": -100..-1 'G_GIF'; 0 'G_PNG'; 1..9 'G_JPG'; 10 'G_BMP'; 32000 'G_SVG'

recipe "Recipe_1": Recipe_element_1 <- "D_Int", Recipe_element_2 <- "D_Real", Recipe_element_3 <- "D_Pct", Recipe_element_4 <- "D_Bits", Recipe_element_5 <- "D_Range"

SlideinScreen "GraphX_Slidein_Top" 1024x120
   TextField "SI_Title" at 10,10 size 127x20; Text 'Slide-in screen Top'
   Bar "SI_Bar" at 330,10 size 200x40
      ProcessValue <- "D_Pct"
   IOField "SI_Value" at 560,10 size 120x30; FormatPattern s99999
      ProcessValue <- "D_Int"

screen "All_Objects" 1024x768
   TextField "TextField_1" at 680,10 size 33x20; Text 'Text'
   GraphicView "GraphicView_1" at 800,10 size 100x60
   IOField "IOField_1" at 10,90 size 100x30
   Button "Button_1" at 130,90 size 100x40; TextOff 'Text'
   SymbolicIOField "SymbolicIOField_1" at 250,90 size 120x30; TextOff '0'; TextOn '1'
   GraphicIOField "GraphicIOField_1" at 390,90 size 60x60
   DateTimeField "DateTimeField_1" at 470,90 size 189x26
   Bar "Bar_1" at 650,90 size 40x120
   Switch "Switch_1" at 710,90 size 120x40; CaptionText 'Switch'; TextOff '0'; TextOn '1'
   SymbolLibrary "SymbolLibrary_1" at 850,90 size 60x60
   Slider "Slider_1" at 930,90 size 60x160; Caption 'SIMATIC'
   Gauge "Gauge_1" at 10,270 size 150x150; CaptionText 'SIMATIC'
   Clock "Clock_1" at 180,270 size 150x150

screen "Ctl_01_AlarmView" 1024x768, template "Nav"
   AlarmView "Alarm view_1" at 3,3 size 600x300

screen "Ctl_02_TrendView" 1024x768, template "Nav"
   TrendView "Trend view_1" at 3,3 size 600x300

screen "Ctl_03_UserView" 1024x768, template "Nav"
   UserView "User view_1" at 3,3 size 480x240

screen "Ctl_04_HtmlBrowser" 1024x768, template "Nav"
   HTMLBrowser "HTML browser_1" at 3,3 size 192x192

screen "Ctl_05_WatchTable" 1024x768, template "Nav"
   StatusForce "Watch table_1" at 3,3 size 600x300; ToolTipText 'Text'

screen "Ctl_06_SmartClientView" 1024x768, template "Nav"
   SmartClientView "Sm@rtClient view_1" at 3,3 size 320x240

screen "Ctl_07_RecipeView" 1024x768, template "Nav"
   RecipeView "Recipe view_1" at 3,3 size 400x330; Recipe "Recipe_1"

screen "Ctl_09_SysDiagView" 1024x768, template "Nav"
   SysDiagControl "System diagnostics view_1" at 3,3 size 600x300

screen "Ctl_10_MediaPlayer" 1024x768, template "Nav"
   MediaPlayer "Media Player_1" at 3,3 size 240x240

screen "Ctl_11_PlcCodeView" 1024x768, template "Nav"
   PLCCodeViewer "PLC code view_1" at 3,3 size 600x300

screen "Ctl_12_GraphOverview" 1024x768, template "Nav"
   S7GraphOverview "GRAPH overview_1" at 3,3 size 424x72

screen "Ctl_13_ProDiagOverview" 1024x768, template "Nav"
   ProDiagOverview "ProDiag overview_1" at 3,3 size 253x72

screen "Ctl_14_CriteriaAnalysisView" 1024x768, template "Nav"
   CriteriaAnalysisView "Criteria analysis view_1" at 3,3 size 460x150

screen "Ctl_15_CameraView" 1024x768, template "Nav"
   CameraControl "Camera view_1" at 3,3 size 320x240

screen "Ctl_16_PdfView" 1024x768, template "Nav"
   PDFView "PDFView_1" at 3,3 size 320x240

Template "Nav" 1024x768
   Button "Nav_01" at 994,2 size 28x22; TextOff 'Text'
      on Click: ActivateScreen("Ctl_01_AlarmView", 0)
   Button "Nav_02" at 994,28 size 28x22; TextOff 'Text'
      on Click: ActivateScreen("Ctl_02_TrendView", 0)
   Button "Nav_03" at 994,54 size 28x22; TextOff 'Text'
      on Click: ActivateScreen("Ctl_03_UserView", 0)
   Button "Nav_04" at 994,80 size 28x22; TextOff 'Text'
      on Click: ActivateScreen("Ctl_04_HtmlBrowser", 0)
   Button "Nav_05" at 994,106 size 28x22; TextOff 'Text'
      on Click: ActivateScreen("Ctl_05_WatchTable", 0)
   Button "Nav_06" at 994,132 size 28x22; TextOff 'Text'
      on Click: ActivateScreen("Ctl_06_SmartClientView", 0)
   Button "Nav_07" at 994,158 size 28x22; TextOff 'Text'
      on Click: ActivateScreen("Ctl_07_RecipeView", 0)
   Button "Nav_09" at 994,210 size 28x22; TextOff 'Text'
      on Click: ActivateScreen("Ctl_09_SysDiagView", 0)
   Button "Nav_10" at 994,236 size 28x22; TextOff 'Text'
      on Click: ActivateScreen("Ctl_10_MediaPlayer", 0)
   Button "Nav_11" at 994,262 size 28x22; TextOff 'Text'
      on Click: ActivateScreen("Ctl_11_PlcCodeView", 0)
   Button "Nav_12" at 994,288 size 28x22; TextOff 'Text'
      on Click: ActivateScreen("Ctl_12_GraphOverview", 0)
   Button "Nav_13" at 994,314 size 28x22; TextOff 'Text'
      on Click: ActivateScreen("Ctl_13_ProDiagOverview", 0)
   Button "Nav_14" at 994,340 size 28x22; TextOff 'Text'
      on Click: ActivateScreen("Ctl_14_CriteriaAnalysisView", 0)
   Button "Nav_15" at 994,366 size 28x22; TextOff 'Text'
      on Click: ActivateScreen("Ctl_15_CameraView", 0)
   Button "Nav_16" at 994,392 size 28x22; TextOff 'Text'
      on Click: ActivateScreen("Ctl_16_PdfView", 0)
   Button "Nav_17" at 994,418 size 28x22; TextOff 'Text'
      on Click: ActivateScreen("All_Objects", 0)

screen "P_Line_1" 1024x768
   TextField "Label_Default" at 10,62 size 52x20; Text 'Default'
   TextField "Label_BackColor" at 120,62 size 68x20; Text 'BackColor'
   TextField "Label_Color" at 230,62 size 38x20; Text 'Color'
   TextField "Label_EndStyle" at 340,62 size 61x20; Text 'EndStyle'
   TextField "Label_EndStyle_2" at 450,62 size 77x20; Text 'EndStyle_2'
   TextField "Label_EndStyle_3" at 560,62 size 77x20; Text 'EndStyle_3'
   TextField "Label_EndStyle_4" at 670,62 size 77x20; Text 'EndStyle_4'
   TextField "Label_EndStyle_5" at 780,62 size 77x20; Text 'EndStyle_5'
   TextField "Label_FillStyle" at 890,62 size 53x20; Text 'FillStyle'
   TextField "Label_Flashing" at 10,138 size 56x20; Text 'Flashing'
   TextField "Label_LineEndShapeStyle_2" at 120,138 size 143x20; Text 'LineEndShapeStyle_2'
   TextField "Label_LineWidth" at 230,138 size 69x20; Text 'LineWidth'
   TextField "Label_StartStyle" at 340,138 size 72x20; Text 'StartStyle'
   TextField "Label_StartStyle_2" at 450,138 size 88x20; Text 'StartStyle_2'
   TextField "Label_StartStyle_3" at 560,138 size 88x20; Text 'StartStyle_3'
   TextField "Label_StartStyle_4" at 670,138 size 88x20; Text 'StartStyle_4'
   TextField "Label_StartStyle_5" at 780,138 size 88x20; Text 'StartStyle_5'
   TextField "Label_Style" at 890,138 size 38x20; Text 'Style'
   TextField "Label_Style_2" at 10,214 size 54x20; Text 'Style_2'
   TextField "Label_Style_3" at 120,214 size 54x20; Text 'Style_3'
   TextField "Label_Style_4" at 230,214 size 54x20; Text 'Style_4'
   TextField "Label_UseDesignColorSchema" at 340,214 size 154x20; Text 'UseDesignColorSchema'
   Button "Next" at 982,744 size 40x22; TextOff 'Text'
      on Click: ActivateScreen("P_Polyline_1", 0)

screen "P_Polyline_1" 1024x768
   TextField "Label_Default" at 10,62 size 52x20; Text 'Default'
   TextField "Label_BackColor" at 120,62 size 68x20; Text 'BackColor'
   TextField "Label_Color" at 230,62 size 38x20; Text 'Color'
   TextField "Label_EndStyle" at 340,62 size 61x20; Text 'EndStyle'
   TextField "Label_EndStyle_2" at 450,62 size 77x20; Text 'EndStyle_2'
   TextField "Label_EndStyle_3" at 560,62 size 77x20; Text 'EndStyle_3'
   TextField "Label_EndStyle_4" at 670,62 size 77x20; Text 'EndStyle_4'
   TextField "Label_EndStyle_5" at 780,62 size 77x20; Text 'EndStyle_5'
   TextField "Label_FillStyle" at 890,62 size 53x20; Text 'FillStyle'
   TextField "Label_Flashing" at 10,138 size 56x20; Text 'Flashing'
   TextField "Label_LineEndShapeStyle_2" at 120,138 size 143x20; Text 'LineEndShapeStyle_2'
   TextField "Label_LineWidth" at 230,138 size 69x20; Text 'LineWidth'
   TextField "Label_StartStyle" at 340,138 size 72x20; Text 'StartStyle'
   TextField "Label_StartStyle_2" at 450,138 size 88x20; Text 'StartStyle_2'
   TextField "Label_StartStyle_3" at 560,138 size 88x20; Text 'StartStyle_3'
   TextField "Label_StartStyle_4" at 670,138 size 88x20; Text 'StartStyle_4'
   TextField "Label_StartStyle_5" at 780,138 size 88x20; Text 'StartStyle_5'
   TextField "Label_Style" at 890,138 size 38x20; Text 'Style'
   TextField "Label_Style_2" at 10,214 size 54x20; Text 'Style_2'
   TextField "Label_Style_3" at 120,214 size 54x20; Text 'Style_3'
   TextField "Label_Style_4" at 230,214 size 54x20; Text 'Style_4'
   TextField "Label_UseDesignColorSchema" at 340,214 size 154x20; Text 'UseDesignColorSchema'
   Button "Next" at 982,744 size 40x22; TextOff 'Text'
      on Click: ActivateScreen("P_Polygon_1", 0)

screen "P_Polygon_1" 1024x768
   TextField "Label_Default" at 10,62 size 52x20; Text 'Default'
   TextField "Label_BackColor" at 120,62 size 68x20; Text 'BackColor'
   TextField "Label_BackFillStyle" at 230,62 size 83x20; Text 'BackFillStyle'
   TextField "Label_BorderColor" at 340,62 size 82x20; Text 'BorderColor'
   TextField "Label_BorderWidth" at 450,62 size 87x20; Text 'BorderWidth'
   TextField "Label_EdgeStyle" at 560,62 size 69x20; Text 'EdgeStyle'
   TextField "Label_EdgeStyle_2" at 670,62 size 85x20; Text 'EdgeStyle_2'
   TextField "Label_EdgeStyle_3" at 780,62 size 85x20; Text 'EdgeStyle_3'
   TextField "Label_EdgeStyle_4" at 890,62 size 85x20; Text 'EdgeStyle_4'
   TextField "Label_Flashing" at 10,138 size 56x20; Text 'Flashing'
   TextField "Label_UseDesignColorSchema" at 120,138 size 154x20; Text 'UseDesignColorSchema'
   Button "Next" at 982,744 size 40x22; TextOff 'Text'
      on Click: ActivateScreen("P_Ellipse_1", 0)

screen "P_Ellipse_1" 1024x768
   TextField "Label_Default" at 10,62 size 52x20; Text 'Default'
   TextField "Label_BackColor" at 120,62 size 68x20; Text 'BackColor'
   TextField "Label_BackFillStyle" at 230,62 size 83x20; Text 'BackFillStyle'
   TextField "Label_BorderColor" at 340,62 size 82x20; Text 'BorderColor'
   TextField "Label_BorderWidth" at 450,62 size 87x20; Text 'BorderWidth'
   TextField "Label_EdgeStyle" at 560,62 size 69x20; Text 'EdgeStyle'
   TextField "Label_EdgeStyle_2" at 670,62 size 85x20; Text 'EdgeStyle_2'
   TextField "Label_EdgeStyle_3" at 780,62 size 85x20; Text 'EdgeStyle_3'
   TextField "Label_EdgeStyle_4" at 890,62 size 85x20; Text 'EdgeStyle_4'
   TextField "Label_Flashing" at 10,138 size 56x20; Text 'Flashing'
   TextField "Label_UseDesignColorSchema" at 120,138 size 154x20; Text 'UseDesignColorSchema'
   Button "Next" at 982,744 size 40x22; TextOff 'Text'
      on Click: ActivateScreen("P_Circle_1", 0)

screen "P_Circle_1" 1024x768
   TextField "Label_Default" at 10,62 size 52x20; Text 'Default'
   TextField "Label_BackColor" at 70,62 size 68x20; Text 'BackColor'
   TextField "Label_BackFillStyle" at 130,62 size 83x20; Text 'BackFillStyle'
   TextField "Label_BorderColor" at 190,62 size 82x20; Text 'BorderColor'
   TextField "Label_BorderWidth" at 250,62 size 87x20; Text 'BorderWidth'
   TextField "Label_EdgeStyle" at 310,62 size 69x20; Text 'EdgeStyle'
   TextField "Label_EdgeStyle_2" at 370,62 size 85x20; Text 'EdgeStyle_2'
   TextField "Label_EdgeStyle_3" at 430,62 size 85x20; Text 'EdgeStyle_3'
   TextField "Label_EdgeStyle_4" at 490,62 size 85x20; Text 'EdgeStyle_4'
   TextField "Label_Flashing" at 550,62 size 56x20; Text 'Flashing'
   TextField "Label_UseDesignColorSchema" at 610,62 size 154x20; Text 'UseDesignColorSchema'
   Button "Next" at 982,744 size 40x22; TextOff 'Text'
      on Click: ActivateScreen("P_Rectangle_1", 0)

screen "P_Rectangle_1" 1024x768
   TextField "Label_Default" at 10,62 size 52x20; Text 'Default'
   TextField "Label_BackColor" at 120,62 size 68x20; Text 'BackColor'
   TextField "Label_BackFillStyle" at 230,62 size 83x20; Text 'BackFillStyle'
   TextField "Label_BorderColor" at 340,62 size 82x20; Text 'BorderColor'
   TextField "Label_BorderWidth" at 450,62 size 87x20; Text 'BorderWidth'
   TextField "Label_EdgeStyle" at 560,62 size 69x20; Text 'EdgeStyle'
   TextField "Label_EdgeStyle_2" at 670,62 size 85x20; Text 'EdgeStyle_2'
   TextField "Label_EdgeStyle_3" at 780,62 size 85x20; Text 'EdgeStyle_3'
   TextField "Label_EdgeStyle_4" at 890,62 size 85x20; Text 'EdgeStyle_4'
   TextField "Label_Flashing" at 10,138 size 56x20; Text 'Flashing'
   TextField "Label_RoundCornerHeight" at 120,138 size 132x20; Text 'RoundCornerHeight'
   TextField "Label_RoundCornerWidth" at 230,138 size 128x20; Text 'RoundCornerWidth'
   TextField "Label_UseDesignColorSchema" at 340,138 size 154x20; Text 'UseDesignColorSchema'
   Button "Next" at 982,744 size 40x22; TextOff 'Text'
      on Click: ActivateScreen("P_TextField_1", 0)

screen "P_TextField_1" 1024x768
   TextField "Default" at 10,10 size 33x20; Text 'Text'
   TextField "Label_Default" at 10,42 size 52x20; Text 'Default'
   TextField "BackColor" at 120,10 size 33x20; Text 'Text'
   TextField "Label_BackColor" at 120,42 size 68x20; Text 'BackColor'
   TextField "BackFillStyle" at 230,10 size 33x20; Text 'Text'
   TextField "Label_BackFillStyle" at 230,42 size 83x20; Text 'BackFillStyle'
   TextField "BorderBackColor" at 340,10 size 33x20; Text 'Text'
   TextField "Label_BorderBackColor" at 340,42 size 112x20; Text 'BorderBackColor'
   TextField "BorderColor" at 450,10 size 33x20; Text 'Text'
   TextField "Label_BorderColor" at 450,42 size 82x20; Text 'BorderColor'
   TextField "BorderWidth" at 560,10 size 33x20; Text 'Text'
   TextField "Label_BorderWidth" at 560,42 size 87x20; Text 'BorderWidth'
   TextField "BottomMargin" at 670,10 size 33x20; Text 'Text'
   TextField "Label_BottomMargin" at 670,42 size 96x20; Text 'BottomMargin'
   TextField "CornerRadius" at 780,10 size 33x20; Text 'Text'
   TextField "Label_CornerRadius" at 780,42 size 92x20; Text 'CornerRadius'
   TextField "EdgeStyle" at 890,10 size 33x20; Text 'Text'
   TextField "Label_EdgeStyle" at 890,42 size 69x20; Text 'EdgeStyle'
   TextField "EdgeStyle_2" at 10,66 size 33x20; Text 'Text'
   TextField "Label_EdgeStyle_2" at 10,98 size 85x20; Text 'EdgeStyle_2'
   TextField "EdgeStyle_3" at 120,66 size 33x20; Text 'Text'
   TextField "Label_EdgeStyle_3" at 120,98 size 85x20; Text 'EdgeStyle_3'
   TextField "EdgeStyle_4" at 230,66 size 33x20; Text 'Text'
   TextField "Label_EdgeStyle_4" at 230,98 size 85x20; Text 'EdgeStyle_4'
   TextField "FitToLargest" at 340,66 size 100x30; Text 'Text'
   TextField "Label_FitToLargest" at 340,98 size 85x20; Text 'FitToLargest'
   TextField "Flashing" at 450,66 size 33x20; Text 'Text'
   TextField "Label_Flashing" at 450,98 size 56x20; Text 'Flashing'
   TextField "ForeColor" at 560,66 size 33x20; Text 'Text'
   TextField "Label_ForeColor" at 560,98 size 66x20; Text 'ForeColor'
   TextField "HorizontalAlignment" at 670,66 size 33x20; Text 'Text'
   TextField "Label_HorizontalAlignment" at 670,98 size 136x20; Text 'HorizontalAlignment'
   TextField "HorizontalAlignment_2" at 780,66 size 33x20; Text 'Text'
   TextField "Label_HorizontalAlignment_2" at 780,98 size 152x20; Text 'HorizontalAlignment_2'
   TextField "LeftMargin" at 890,66 size 33x20; Text 'Text'
   TextField "Label_LeftMargin" at 890,98 size 75x20; Text 'LeftMargin'
   TextField "RightMargin" at 10,122 size 33x20; Text 'Text'
   TextField "Label_RightMargin" at 10,154 size 83x20; Text 'RightMargin'
   TextField "TopMargin" at 120,122 size 33x20; Text 'Text'
   TextField "Label_TopMargin" at 120,154 size 72x20; Text 'TopMargin'
   TextField "UseDesignColorSchema" at 230,122 size 33x21; Text 'Text'
   TextField "Label_UseDesignColorSchema" at 230,154 size 154x20; Text 'UseDesignColorSchema'
   TextField "VerticalAlignment" at 340,122 size 33x20; Text 'Text'
   TextField "Label_VerticalAlignment" at 340,154 size 120x20; Text 'VerticalAlignment'
   TextField "VerticalAlignment_2" at 450,122 size 33x20; Text 'Text'
   TextField "Label_VerticalAlignment_2" at 450,154 size 136x20; Text 'VerticalAlignment_2'
   Button "Next" at 982,744 size 40x22; TextOff 'Text'
      on Click: ActivateScreen("P_GraphicView_1", 0)

screen "P_GraphicView_1" 1024x768
   GraphicView "Default" at 10,10 size 100x60
   TextField "Label_Default" at 10,72 size 52x20; Text 'Default'
   GraphicView "BackColor" at 120,10 size 100x60
   TextField "Label_BackColor" at 120,72 size 68x20; Text 'BackColor'
   GraphicView "BackFillStyle" at 230,10 size 100x60
   TextField "Label_BackFillStyle" at 230,72 size 83x20; Text 'BackFillStyle'
   GraphicView "BorderColor" at 340,10 size 100x60
   TextField "Label_BorderColor" at 340,72 size 82x20; Text 'BorderColor'
   GraphicView "BorderWidth" at 450,10 size 100x60
   TextField "Label_BorderWidth" at 450,72 size 87x20; Text 'BorderWidth'
   GraphicView "EdgeStyle" at 560,10 size 100x60
   TextField "Label_EdgeStyle" at 560,72 size 69x20; Text 'EdgeStyle'
   GraphicView "EdgeStyle_2" at 670,10 size 100x60
   TextField "Label_EdgeStyle_2" at 670,72 size 85x20; Text 'EdgeStyle_2'
   GraphicView "EdgeStyle_3" at 780,10 size 100x60
   TextField "Label_EdgeStyle_3" at 780,72 size 85x20; Text 'EdgeStyle_3'
   GraphicView "EdgeStyle_4" at 890,10 size 100x60
   TextField "Label_EdgeStyle_4" at 890,72 size 85x20; Text 'EdgeStyle_4'
   GraphicView "FitToLargest" at 10,96 size 100x60
   TextField "Label_FitToLargest" at 10,158 size 85x20; Text 'FitToLargest'
   GraphicView "Flashing" at 120,96 size 100x60
   TextField "Label_Flashing" at 120,158 size 56x20; Text 'Flashing'
   GraphicView "TransparentColor" at 230,96 size 100x60
   TextField "Label_TransparentColor" at 230,158 size 118x20; Text 'TransparentColor'
   GraphicView "UseTransparentColor" at 340,96 size 100x60
   TextField "Label_UseTransparentColor" at 340,158 size 141x20; Text 'UseTransparentColor'
   Button "Next" at 982,744 size 40x22; TextOff 'Text'
      on Click: ActivateScreen("P_IOField_1", 0)

screen "P_Button_1" 1024x768
   Button "Default" at 10,10 size 100x40; TextOff 'Text'
   TextField "Label_Default" at 10,52 size 52x20; Text 'Default'
   Button "BackColor" at 120,10 size 100x40; TextOff 'Text'
   TextField "Label_BackColor" at 120,52 size 68x20; Text 'BackColor'
   Button "BackFillStyle" at 230,10 size 100x40; TextOff 'Text'
   TextField "Label_BackFillStyle" at 230,52 size 83x20; Text 'BackFillStyle'
   Button "BorderBackColor" at 340,10 size 100x40; TextOff 'Text'
   TextField "Label_BorderBackColor" at 340,52 size 112x20; Text 'BorderBackColor'
   Button "BorderColor" at 450,10 size 100x40; TextOff 'Text'
   TextField "Label_BorderColor" at 450,52 size 82x20; Text 'BorderColor'
   Button "BorderWidth" at 560,10 size 100x40; TextOff 'Text'
   TextField "Label_BorderWidth" at 560,52 size 87x20; Text 'BorderWidth'
   Button "CornerRadius" at 670,10 size 100x40; TextOff 'Text'
   TextField "Label_CornerRadius" at 670,52 size 92x20; Text 'CornerRadius'
   Button "EdgeStyle" at 780,10 size 100x40; TextOff 'Text'
   TextField "Label_EdgeStyle" at 780,52 size 69x20; Text 'EdgeStyle'
   Button "EdgeStyle_2" at 890,10 size 100x40; TextOff 'Text'
   TextField "Label_EdgeStyle_2" at 890,52 size 85x20; Text 'EdgeStyle_2'
   Button "EdgeStyle_3" at 10,76 size 100x40; TextOff 'Text'
   TextField "Label_EdgeStyle_3" at 10,118 size 85x20; Text 'EdgeStyle_3'
   Button "EdgeStyle_4" at 120,76 size 100x40; TextOff 'Text'
   TextField "Label_EdgeStyle_4" at 120,118 size 85x20; Text 'EdgeStyle_4'
   Button "FirstGradientColor" at 230,76 size 100x40; TextOff 'Text'
   TextField "Label_FirstGradientColor" at 230,118 size 121x20; Text 'FirstGradientColor'
   Button "FirstGradientOffset" at 340,76 size 100x40; TextOff 'Text'
   TextField "Label_FirstGradientOffset" at 340,118 size 128x20; Text 'FirstGradientOffset'
   Button "FitToLargest" at 450,76 size 32x23; TextOff 'Text'
   TextField "Label_FitToLargest" at 450,118 size 85x20; Text 'FitToLargest'
   Button "Flashing" at 560,76 size 100x40; TextOff 'Text'
   TextField "Label_Flashing" at 560,118 size 56x20; Text 'Flashing'
   Button "FocusColor" at 670,76 size 100x40; TextOff 'Text'
   TextField "Label_FocusColor" at 670,118 size 74x20; Text 'FocusColor'
   Button "FocusWidth" at 780,76 size 100x40; TextOff 'Text'
   TextField "Label_FocusWidth" at 780,118 size 79x20; Text 'FocusWidth'
   Button "ForeColor" at 890,76 size 100x40; TextOff 'Text'
   TextField "Label_ForeColor" at 890,118 size 66x20; Text 'ForeColor'
   Button "HorizontalAlignment" at 10,142 size 100x40; TextOff 'Text'
   TextField "Label_HorizontalAlignment" at 10,184 size 136x20; Text 'HorizontalAlignment'
   Button "HorizontalAlignment_2" at 120,142 size 100x40; TextOff 'Text'
   TextField "Label_HorizontalAlignment_2" at 120,184 size 152x20; Text 'HorizontalAlignment_2'
   Button "HorizontalPictureAlignment" at 230,142 size 100x40; TextOff 'Text'
   TextField "Label_HorizontalPictureAlignment" at 230,184 size 182x20; Text 'HorizontalPictureAlignment'
   Button "HorizontalPictureAlignment_2" at 340,142 size 100x40; TextOff 'Text'
   TextField "Label_HorizontalPictureAlignment_2" at 340,184 size 198x20; Text 'HorizontalPictureAlignment_2'
   Button "MiddleGradientColor" at 450,142 size 100x40; TextOff 'Text'
   TextField "Label_MiddleGradientColor" at 450,184 size 134x20; Text 'MiddleGradientColor'
   Button "Mode_5" at 560,142 size 100x40; TextOff 'Text'
   TextField "Label_Mode_5" at 560,184 size 56x20; Text 'Mode_5'
   Button "Mode_7" at 670,142 size 100x40; TextOff 'Text'
   TextField "Label_Mode_7" at 670,184 size 56x20; Text 'Mode_7'
   Button "PictureAreaBottomMargin" at 780,142 size 100x40; TextOff 'Text'
   TextField "Label_PictureAreaBottomMargin" at 780,184 size 174x20; Text 'PictureAreaBottomMargin'
   Button "PictureAreaLeftMargin" at 890,142 size 100x40; TextOff 'Text'
   TextField "Label_PictureAreaLeftMargin" at 890,184 size 153x20; Text 'PictureAreaLeftMargin'
   Button "PictureAreaRightMargin" at 10,208 size 100x40; TextOff 'Text'
   TextField "Label_PictureAreaRightMargin" at 10,250 size 161x20; Text 'PictureAreaRightMargin'
   Button "PictureAreaTopMargin" at 120,208 size 100x40; TextOff 'Text'
   TextField "Label_PictureAreaTopMargin" at 120,250 size 150x20; Text 'PictureAreaTopMargin'
   Button "SecondGradientColor" at 230,208 size 100x40; TextOff 'Text'
   TextField "Label_SecondGradientColor" at 230,250 size 140x20; Text 'SecondGradientColor'
   Button "SecondGradientOffset" at 340,208 size 100x40; TextOff 'Text'
   TextField "Label_SecondGradientOffset" at 340,250 size 147x20; Text 'SecondGradientOffset'
   Button "TextAreaBottomMargin" at 450,208 size 100x40; TextOff 'Text'
   TextField "Label_TextAreaBottomMargin" at 450,250 size 156x20; Text 'TextAreaBottomMargin'
   Button "TextAreaLeftMargin" at 560,208 size 100x40; TextOff 'Text'
   TextField "Label_TextAreaLeftMargin" at 560,250 size 135x20; Text 'TextAreaLeftMargin'
   Button "TextAreaRightMargin" at 670,208 size 100x40; TextOff 'Text'
   TextField "Label_TextAreaRightMargin" at 670,250 size 143x20; Text 'TextAreaRightMargin'
   Button "TextAreaTopMargin" at 780,208 size 100x40; TextOff 'Text'
   TextField "Label_TextAreaTopMargin" at 780,250 size 132x20; Text 'TextAreaTopMargin'
   Button "UseDesignColorSchema" at 890,208 size 100x40; TextOff 'Text'
   TextField "Label_UseDesignColorSchema" at 890,250 size 154x20; Text 'UseDesignColorSchema'
   Button "UseFirstGradient" at 10,274 size 100x40; TextOff 'Text'
   TextField "Label_UseFirstGradient" at 10,316 size 111x20; Text 'UseFirstGradient'
   Button "UseSecondGradient" at 120,274 size 100x40; TextOff 'Text'
   TextField "Label_UseSecondGradient" at 120,316 size 130x20; Text 'UseSecondGradient'
   Button "VerticalAlignment" at 230,274 size 100x40; TextOff 'Text'
   TextField "Label_VerticalAlignment" at 230,316 size 120x20; Text 'VerticalAlignment'
   Button "VerticalAlignment_2" at 340,274 size 100x40; TextOff 'Text'
   TextField "Label_VerticalAlignment_2" at 340,316 size 136x20; Text 'VerticalAlignment_2'
   Button "VerticalPictureAlignment" at 450,274 size 100x40; TextOff 'Text'
   TextField "Label_VerticalPictureAlignment" at 450,316 size 166x20; Text 'VerticalPictureAlignment'
   Button "VerticalPictureAlignment_2" at 560,274 size 100x40; TextOff 'Text'
   TextField "Label_VerticalPictureAlignment_2" at 560,316 size 182x20; Text 'VerticalPictureAlignment_2'
   Button "Next" at 982,744 size 40x22; TextOff 'Text'
      on Click: ActivateScreen("P_SymbolicIOField_1", 0)

screen "P_SymbolicIOField_1" 1024x768
   SymbolicIOField "Default" at 10,10 size 120x30; TextOff '0'; TextOn '1'
   TextField "Label_Default" at 10,42 size 52x20; Text 'Default'
   SymbolicIOField "AboveUpperLimitColor" at 140,10 size 120x30; TextOff '0'; TextOn '1'
   TextField "Label_AboveUpperLimitColor" at 140,42 size 148x20; Text 'AboveUpperLimitColor'
   SymbolicIOField "BackColor" at 270,10 size 120x30; TextOff '0'; TextOn '1'
   TextField "Label_BackColor" at 270,42 size 68x20; Text 'BackColor'
   SymbolicIOField "BackFillStyle" at 400,10 size 120x30; TextOff '0'; TextOn '1'
   TextField "Label_BackFillStyle" at 400,42 size 83x20; Text 'BackFillStyle'
   SymbolicIOField "BelowLowerLimitColor" at 530,10 size 120x30; TextOff '0'; TextOn '1'
   TextField "Label_BelowLowerLimitColor" at 530,42 size 146x20; Text 'BelowLowerLimitColor'
   SymbolicIOField "BorderBackColor" at 660,10 size 120x30; TextOff '0'; TextOn '1'
   TextField "Label_BorderBackColor" at 660,42 size 112x20; Text 'BorderBackColor'
   SymbolicIOField "BorderColor" at 790,10 size 120x30; TextOff '0'; TextOn '1'
   TextField "Label_BorderColor" at 790,42 size 82x20; Text 'BorderColor'
   SymbolicIOField "BorderWidth" at 10,66 size 120x30; TextOff '0'; TextOn '1'
   TextField "Label_BorderWidth" at 10,98 size 87x20; Text 'BorderWidth'
   SymbolicIOField "BottomMargin" at 140,66 size 120x30; TextOff '0'; TextOn '1'
   TextField "Label_BottomMargin" at 140,98 size 96x20; Text 'BottomMargin'
   SymbolicIOField "CornerRadius" at 270,66 size 120x30; TextOff '0'; TextOn '1'
   TextField "Label_CornerRadius" at 270,98 size 92x20; Text 'CornerRadius'
   SymbolicIOField "CountVisibleItems" at 400,66 size 120x30; TextOff '0'; TextOn '1'
   TextField "Label_CountVisibleItems" at 400,98 size 121x20; Text 'CountVisibleItems'
   SymbolicIOField "EdgeStyle" at 530,66 size 120x30; TextOff '0'; TextOn '1'
   TextField "Label_EdgeStyle" at 530,98 size 69x20; Text 'EdgeStyle'
   SymbolicIOField "EdgeStyle_2" at 660,66 size 120x30; TextOff '0'; TextOn '1'
   TextField "Label_EdgeStyle_2" at 660,98 size 85x20; Text 'EdgeStyle_2'
   SymbolicIOField "EdgeStyle_3" at 790,66 size 120x30; TextOff '0'; TextOn '1'
   TextField "Label_EdgeStyle_3" at 790,98 size 85x20; Text 'EdgeStyle_3'
   SymbolicIOField "EdgeStyle_4" at 10,122 size 120x30; TextOff '0'; TextOn '1'
   TextField "Label_EdgeStyle_4" at 10,154 size 85x20; Text 'EdgeStyle_4'
   SymbolicIOField "EvenRowBackColor" at 140,122 size 120x30; TextOff '0'; TextOn '1'
   TextField "Label_EvenRowBackColor" at 140,154 size 127x20; Text 'EvenRowBackColor'
   SymbolicIOField "FitToLargest" at 270,122 size 41x28; TextOff '0'; TextOn '1'
   TextField "Label_FitToLargest" at 270,154 size 85x20; Text 'FitToLargest'
   SymbolicIOField "Flashing" at 400,122 size 120x30; TextOff '0'; TextOn '1'
   TextField "Label_Flashing" at 400,154 size 56x20; Text 'Flashing'
   SymbolicIOField "FlashingOnLimitViolation" at 530,122 size 120x30; TextOff '0'; TextOn '1'
   TextField "Label_FlashingOnLimitViolation" at 530,154 size 159x20; Text 'FlashingOnLimitViolation'
   SymbolicIOField "ForeColor" at 660,122 size 120x30; TextOff '0'; TextOn '1'
   TextField "Label_ForeColor" at 660,154 size 66x20; Text 'ForeColor'
   SymbolicIOField "HorizontalAlignment" at 790,122 size 120x30; TextOff '0'; TextOn '1'
   TextField "Label_HorizontalAlignment" at 790,154 size 136x20; Text 'HorizontalAlignment'
   SymbolicIOField "HorizontalAlignment_2" at 10,178 size 120x30; TextOff '0'; TextOn '1'
   TextField "Label_HorizontalAlignment_2" at 10,210 size 152x20; Text 'HorizontalAlignment_2'
   SymbolicIOField "LeftMargin" at 140,178 size 120x30; TextOff '0'; TextOn '1'
   TextField "Label_LeftMargin" at 140,210 size 75x20; Text 'LeftMargin'
   SymbolicIOField "Mode" at 270,178 size 120x30; TextOff '0'; TextOn '1'
   TextField "Label_Mode" at 270,210 size 40x20; Text 'Mode'
   SymbolicIOField "Mode_2" at 400,178 size 120x30; TextOff '0'; TextOn '1'
   TextField "Label_Mode_2" at 400,210 size 56x20; Text 'Mode_2'
   SymbolicIOField "RightMargin" at 530,178 size 120x30; TextOff '0'; TextOn '1'
   TextField "Label_RightMargin" at 530,210 size 83x20; Text 'RightMargin'
   SymbolicIOField "SelectBackColor" at 660,178 size 120x30; TextOff '0'; TextOn '1'
   TextField "Label_SelectBackColor" at 660,210 size 108x20; Text 'SelectBackColor'
   SymbolicIOField "SelectForeColor" at 790,178 size 120x30; TextOff '0'; TextOn '1'
   TextField "Label_SelectForeColor" at 790,210 size 106x20; Text 'SelectForeColor'
   SymbolicIOField "ShowDropDownButton" at 10,234 size 120x30; TextOff '0'; TextOn '1'
   TextField "Label_ShowDropDownButton" at 10,266 size 151x20; Text 'ShowDropDownButton'
   SymbolicIOField "ShowDropDownList" at 140,234 size 120x30; TextOff '0'; TextOn '1'
   TextField "Label_ShowDropDownList" at 140,266 size 130x20; Text 'ShowDropDownList'
   SymbolicIOField "TopMargin" at 270,234 size 120x30; TextOff '0'; TextOn '1'
   TextField "Label_TopMargin" at 270,266 size 72x20; Text 'TopMargin'
   SymbolicIOField "UseDesignColorSchema" at 400,234 size 120x30; TextOff '0'; TextOn '1'
   TextField "Label_UseDesignColorSchema" at 400,266 size 154x20; Text 'UseDesignColorSchema'
   SymbolicIOField "VerticalAlignment" at 530,234 size 120x30; TextOff '0'; TextOn '1'
   TextField "Label_VerticalAlignment" at 530,266 size 120x20; Text 'VerticalAlignment'
   SymbolicIOField "VerticalAlignment_2" at 660,234 size 120x30; TextOff '0'; TextOn '1'
   TextField "Label_VerticalAlignment_2" at 660,266 size 136x20; Text 'VerticalAlignment_2'
   Button "Next" at 982,744 size 40x22; TextOff 'Text'
      on Click: ActivateScreen("P_GraphicIOField_1", 0)

screen "P_GraphicIOField_1" 1024x768
   GraphicIOField "Default" at 10,10 size 60x60
   TextField "Label_Default" at 10,72 size 52x20; Text 'Default'
   GraphicIOField "AboveUpperLimitColor" at 80,10 size 60x60
   TextField "Label_AboveUpperLimitColor" at 80,72 size 148x20; Text 'AboveUpperLimitColor'
   GraphicIOField "BackColor" at 150,10 size 60x60
   TextField "Label_BackColor" at 150,72 size 68x20; Text 'BackColor'
   GraphicIOField "BackFillStyle" at 220,10 size 60x60
   TextField "Label_BackFillStyle" at 220,72 size 83x20; Text 'BackFillStyle'
   GraphicIOField "BelowLowerLimitColor" at 290,10 size 60x60
   TextField "Label_BelowLowerLimitColor" at 290,72 size 146x20; Text 'BelowLowerLimitColor'
   GraphicIOField "BorderColor" at 360,10 size 60x60
   TextField "Label_BorderColor" at 360,72 size 82x20; Text 'BorderColor'
   GraphicIOField "BorderWidth" at 430,10 size 60x60
   TextField "Label_BorderWidth" at 430,72 size 87x20; Text 'BorderWidth'
   GraphicIOField "EdgeStyle" at 500,10 size 60x60
   TextField "Label_EdgeStyle" at 500,72 size 69x20; Text 'EdgeStyle'
   GraphicIOField "EdgeStyle_2" at 570,10 size 60x60
   TextField "Label_EdgeStyle_2" at 570,72 size 85x20; Text 'EdgeStyle_2'
   GraphicIOField "EdgeStyle_3" at 640,10 size 60x60
   TextField "Label_EdgeStyle_3" at 640,72 size 85x20; Text 'EdgeStyle_3'
   GraphicIOField "EdgeStyle_4" at 710,10 size 60x60
   TextField "Label_EdgeStyle_4" at 710,72 size 85x20; Text 'EdgeStyle_4'
   GraphicIOField "FitToLargest" at 780,10 size 60x60
   TextField "Label_FitToLargest" at 780,72 size 85x20; Text 'FitToLargest'
   GraphicIOField "Flashing" at 850,10 size 60x60
   TextField "Label_Flashing" at 850,72 size 56x20; Text 'Flashing'
   GraphicIOField "FlashingOnLimitViolation" at 920,10 size 60x60
   TextField "Label_FlashingOnLimitViolation" at 920,72 size 159x20; Text 'FlashingOnLimitViolation'
   GraphicIOField "FocusColor" at 10,96 size 60x60
   TextField "Label_FocusColor" at 10,158 size 74x20; Text 'FocusColor'
   GraphicIOField "FocusWidth" at 80,96 size 60x60
   TextField "Label_FocusWidth" at 80,158 size 79x20; Text 'FocusWidth'
   GraphicIOField "Mode" at 150,96 size 60x60
   TextField "Label_Mode" at 150,158 size 40x20; Text 'Mode'
   GraphicIOField "Mode_2" at 220,96 size 60x60
   TextField "Label_Mode_2" at 220,158 size 56x20; Text 'Mode_2'
   GraphicIOField "ScrollBarOrientation" at 290,96 size 60x60
   TextField "Label_ScrollBarOrientation" at 290,158 size 135x20; Text 'ScrollBarOrientation'
   GraphicIOField "TransparentColor" at 360,96 size 60x60
   TextField "Label_TransparentColor" at 360,158 size 118x20; Text 'TransparentColor'
   GraphicIOField "UseTransparentColor" at 430,96 size 60x60
   TextField "Label_UseTransparentColor" at 430,158 size 141x20; Text 'UseTransparentColor'
   Button "Next" at 982,744 size 40x22; TextOff 'Text'
      on Click: ActivateScreen("P_DateTimeField_1", 0)

screen "P_DateTimeField_1" 1024x768
   DateTimeField "Default" at 10,10 size 189x26
   TextField "Label_Default" at 10,42 size 52x20; Text 'Default'
   DateTimeField "BackColor" at 180,10 size 189x26
   TextField "Label_BackColor" at 180,42 size 68x20; Text 'BackColor'
   DateTimeField "BackFillStyle" at 350,10 size 189x26
   TextField "Label_BackFillStyle" at 350,42 size 83x20; Text 'BackFillStyle'
   DateTimeField "BorderBackColor" at 520,10 size 189x26
   TextField "Label_BorderBackColor" at 520,42 size 112x20; Text 'BorderBackColor'
   DateTimeField "BorderColor" at 690,10 size 189x26
   TextField "Label_BorderColor" at 690,42 size 82x20; Text 'BorderColor'
   DateTimeField "BorderWidth" at 10,66 size 195x32
   TextField "Label_BorderWidth" at 10,98 size 87x20; Text 'BorderWidth'
   DateTimeField "BottomMargin" at 180,66 size 189x32
   TextField "Label_BottomMargin" at 180,98 size 96x20; Text 'BottomMargin'
   DateTimeField "CornerRadius" at 350,66 size 189x26
   TextField "Label_CornerRadius" at 350,98 size 92x20; Text 'CornerRadius'
   DateTimeField "DisplaySystemTime" at 520,66 size 189x26
   TextField "Label_DisplaySystemTime" at 520,98 size 128x20; Text 'DisplaySystemTime'
   DateTimeField "EdgeStyle" at 690,66 size 189x26
   TextField "Label_EdgeStyle" at 690,98 size 69x20; Text 'EdgeStyle'
   DateTimeField "EdgeStyle_2" at 10,122 size 189x26
   TextField "Label_EdgeStyle_2" at 10,154 size 85x20; Text 'EdgeStyle_2'
   DateTimeField "EdgeStyle_3" at 180,122 size 189x26
   TextField "Label_EdgeStyle_3" at 180,154 size 85x20; Text 'EdgeStyle_3'
   DateTimeField "EdgeStyle_4" at 350,122 size 189x26
   TextField "Label_EdgeStyle_4" at 350,154 size 85x20; Text 'EdgeStyle_4'
   DateTimeField "FitToLargest" at 520,122 size 160x30
   TextField "Label_FitToLargest" at 520,154 size 85x20; Text 'FitToLargest'
   DateTimeField "Flashing" at 690,122 size 189x26
   TextField "Label_Flashing" at 690,154 size 56x20; Text 'Flashing'
   DateTimeField "ForeColor" at 10,178 size 189x26
   TextField "Label_ForeColor" at 10,210 size 66x20; Text 'ForeColor'
   DateTimeField "HorizontalAlignment" at 180,178 size 189x26
   TextField "Label_HorizontalAlignment" at 180,210 size 136x20; Text 'HorizontalAlignment'
   DateTimeField "HorizontalAlignment_2" at 350,178 size 189x26
   TextField "Label_HorizontalAlignment_2" at 350,210 size 152x20; Text 'HorizontalAlignment_2'
   DateTimeField "LeftMargin" at 520,178 size 195x26
   TextField "Label_LeftMargin" at 520,210 size 75x20; Text 'LeftMargin'
   DateTimeField "LongDateTimeFormat" at 690,178 size 340x26
   TextField "Label_LongDateTimeFormat" at 690,210 size 141x20; Text 'LongDateTimeFormat'
   DateTimeField "Mode_3" at 10,234 size 189x26
   TextField "Label_Mode_3" at 10,266 size 56x20; Text 'Mode_3'
   DateTimeField "RightMargin" at 180,234 size 195x26
   TextField "Label_RightMargin" at 180,266 size 83x20; Text 'RightMargin'
   DateTimeField "ShowDate" at 350,234 size 100x26
   TextField "Label_ShowDate" at 350,266 size 71x20; Text 'ShowDate'
   DateTimeField "ShowTime" at 520,234 size 90x26
   TextField "Label_ShowTime" at 520,266 size 69x20; Text 'ShowTime'
   DateTimeField "TopMargin" at 690,234 size 189x32
   TextField "Label_TopMargin" at 690,266 size 72x20; Text 'TopMargin'
   DateTimeField "UseDesignColorSchema" at 10,290 size 180x29
   TextField "Label_UseDesignColorSchema" at 10,322 size 154x20; Text 'UseDesignColorSchema'
   DateTimeField "VerticalAlignment" at 180,290 size 189x26
   TextField "Label_VerticalAlignment" at 180,322 size 120x20; Text 'VerticalAlignment'
   DateTimeField "VerticalAlignment_2" at 350,290 size 189x26
   TextField "Label_VerticalAlignment_2" at 350,322 size 136x20; Text 'VerticalAlignment_2'
   Button "Next" at 982,744 size 40x22; TextOff 'Text'
      on Click: ActivateScreen("P_Bar_1", 0)

